TYPE "Sensor Check Struct"
VERSION : 0.1


  STRUCT
   Rising_Pulse_1 : BOOL ;
   Rising_Pulse_2 : BOOL ;
   Memory_Bit_1 : BOOL ;
   Memory_Bit_2 : BOOL ;
   Word_buffer : INT ;
   Word_Result : INT ;
  END_STRUCT ;
END_TYPE

TYPE "CounterCmd"


  STRUCT
   JOB_WR : STRUCT 	// write commands
    NO : BYTE ;	// number
    BUSY : BOOL ;	// job in working
    DONE : BOOL ;	// job is done
    IMPOSS : BOOL ;	// job impossible
    UNKOWN : BOOL ;	// job unkown
   END_STRUCT ;
   JOB_RD : STRUCT 	// read commands
    NO : BYTE ;	// number
    BUSY : BOOL ;	// job in working
    DONE : BOOL ;	// job is done
    IMPOSS : BOOL ;	// job impossible
    UNKOWN : BOOL ;	// job unkown
   END_STRUCT ;
   RESERV_0 : ARRAY  [1 .. 3 ] OF WORD  := 3 (W#16#0) ;	// reserved
   RESERV_1 : WORD ;	// reserved
   MOD_ADR : WORD ;	// module address
   CH_ADR : DWORD ;	// channel address
   DS_OFFS : BYTE ;	// data block offset
   RESERV_2 : BYTE ;	// reserved
   CONTROL_SIGNALS : STRUCT 	// control signals
    BIT0_0 : BOOL ;	// reserved
    BIT0_1 : BOOL ;	// reserved
    BIT0_2 : BOOL ;	// reserved
    BIT0_3 : BOOL ;	// reserved
    BIT0_4 : BOOL ;	// reserved
    BIT0_5 : BOOL ;	// reserved
    BIT0_6 : BOOL ;	// reserved
    BIT0_7 : BOOL ;	// reserved
    CTRL_DQ0 : BOOL ;	// control digital output DQ0
    CTRL_DQ1 : BOOL ;	// control digital output DQ1
    CTRL_DQ2 : BOOL ;	// control digital output DQ2
    CTRL_DQ3 : BOOL ;	// control digital output DQ3
    CTRL_DQ4 : BOOL ;	// control digital output DQ4
    CTRL_DQ5 : BOOL ;	// control digital output DQ5
    CTRL_DQ6 : BOOL ;	// control digital output DQ6
    CTRL_DQ7 : BOOL ;	// control digital output DQ7
    SET_DQ0 : BOOL ;	// set digital output DQ0
    SET_DQ1 : BOOL ;	// set digital output DQ1
    SET_DQ2 : BOOL ;	// set digital output DQ2
    SET_DQ3 : BOOL ;	// set digital output DQ3
    SET_DQ4 : BOOL ;	// set digital output DQ4
    SET_DQ5 : BOOL ;	// set digital output DQ5
    SET_DQ6 : BOOL ;	// set digital output DQ6
    SET_DQ7 : BOOL ;	// set digital output DQ7
    SW_GATE0 : BOOL ;	// software gate 0
    SW_GATE1 : BOOL ;	// software gate 1
    SW_GATE2 : BOOL ;	// software gate 2
    SW_GATE3 : BOOL ;	// software gate 3
    SW_GATE4 : BOOL ;	// software gate 4
    SW_GATE5 : BOOL ;	// software gate 5
    SW_GATE6 : BOOL ;	// software gate 6
    SW_GATE7 : BOOL ;	// software gate 7
    CTRL_DWORD1 : DWORD ;	// reserved
    CTRL_DWORD2 : DWORD ;	// reserved
    CTRL_DWORD3 : DWORD ;	// reserved
   END_STRUCT ;
   CHECKBACK_SIGNALS : STRUCT 	// checkback signals
    BIT0_0 : BOOL ;	// reserved
    STS_TFB : BOOL ;	// status test free bit
    BIT0_2 : BOOL ;	// reserved
    BIT0_3 : BOOL ;	// reserved
    DATA_ERR : BOOL ;	// data error bit
    BIT0_5 : BOOL ;	// reserved
    BIT0_6 : BOOL ;	// reserved
    PARA : BOOL ;	// module parametrized
    STS_CMP0 : BOOL ;	// status compare event 0
    STS_CMP1 : BOOL ;	// status compare event 1
    STS_CMP2 : BOOL ;	// status compare event 2
    STS_CMP3 : BOOL ;	// status compare event 3
    STS_CMP4 : BOOL ;	// status compare event 4
    STS_CMP5 : BOOL ;	// status compare event 5
    STS_CMP6 : BOOL ;	// status compare event 6
    STS_CMP7 : BOOL ;	// status compare event 7
    STS_UFLW0 : BOOL ;	// status counter 0 passed the underflow value
    STS_UFLW1 : BOOL ;	// status counter 1 passed the underflow value
    STS_UFLW2 : BOOL ;	// status counter 2 passed the underflow value
    STS_UFLW3 : BOOL ;	// status counter 3 passed the underflow value
    STS_UFLW4 : BOOL ;	// status counter 4 passed the underflow value
    STS_UFLW5 : BOOL ;	// status counter 5 passed the underflow value
    STS_UFLW6 : BOOL ;	// status counter 6 passed the underflow value
    STS_UFLW7 : BOOL ;	// status counter 7 passed the underflow value
    STS_OFLW0 : BOOL ;	// status counter 0 passed the overflow value
    STS_OFLW1 : BOOL ;	// status counter 1 passed the overflow value
    STS_OFLW2 : BOOL ;	// status counter 2 passed the overflow value
    STS_OFLW3 : BOOL ;	// status counter 3 passed the overflow value
    STS_OFLW4 : BOOL ;	// status counter 4 passed the overflow value
    STS_OFLW5 : BOOL ;	// status counter 5 passed the overflow value
    STS_OFLW6 : BOOL ;	// status counter 6 passed the overflow value
    STS_OFLW7 : BOOL ;	// status counter 7 passed the overflow value
    STS_DIR0 : BOOL ;	// status counter 0 direction
    STS_DIR1 : BOOL ;	// status counter 1 direction
    STS_DIR2 : BOOL ;	// status counter 2 direction
    STS_DIR3 : BOOL ;	// status counter 3 direction
    STS_DIR4 : BOOL ;	// status counter 4 direction
    STS_DIR5 : BOOL ;	// status counter 5 direction
    STS_DIR6 : BOOL ;	// status counter 6 direction
    STS_DIR7 : BOOL ;	// status counter 7 direction
    STS_DI0 : BOOL ;	// status of the digital input 0
    STS_DI1 : BOOL ;	// status of the digital input 1
    STS_DI2 : BOOL ;	// status of the digital input 2
    STS_DI3 : BOOL ;	// status of the digital input 3
    STS_DI4 : BOOL ;	// status of the digital input 4
    STS_DI5 : BOOL ;	// status of the digital input 5
    STS_DI6 : BOOL ;	// status of the digital input 6
    STS_DI7 : BOOL ;	// status of the digital input 7
    STS_DQ0 : BOOL ;	// status of the digital output 0
    STS_DQ1 : BOOL ;	// status of the digital output 1
    STS_DQ2 : BOOL ;	// status of the digital output 2
    STS_DQ3 : BOOL ;	// status of the digital output 3
    STS_DQ4 : BOOL ;	// status of the digital output 4
    STS_DQ5 : BOOL ;	// status of the digital output 5
    STS_DQ6 : BOOL ;	// status of the digital output 6
    STS_DQ7 : BOOL ;	// status of the digital output 7
    STS_GATE0 : BOOL ;	// status of the internal gate 0
    STS_GATE1 : BOOL ;	// status of the internal gate 1
    STS_GATE2 : BOOL ;	// status of the internal gate 2
    STS_GATE3 : BOOL ;	// status of the internal gate 3
    STS_GATE4 : BOOL ;	// status of the internal gate 4
    STS_GATE5 : BOOL ;	// status of the internal gate 5
    STS_GATE6 : BOOL ;	// status of the internal gate 6
    STS_GATE7 : BOOL ;	// status of the internal gate 7
    USER_STAT_WORD0 : WORD ;	// user specific status
    USER_STAT_WORD1 : WORD ;	// user specific status
    USER_STAT_WORD2 : WORD ;	// user specific status
    USER_STAT_WORD3 : WORD ;	// user specific status
   END_STRUCT ;
   LOAD_VAL0 : DINT ;	// load value counter 0
   LOAD_VAL1 : DINT ;	// load value counter 1
   LOAD_VAL2 : DINT ;	// load value counter 2
   LOAD_VAL3 : DINT ;	// load value counter 3
   LOAD_VAL4 : DINT ;	// load value counter 4
   LOAD_VAL5 : DINT ;	// load value counter 5
   LOAD_VAL6 : DINT ;	// load value counter 6
   LOAD_VAL7 : DINT ;	// load value counter 7
   LOAD_PREPARE_VAL0 : DINT ;	// load prepare value counter 0
   LOAD_PREPARE_VAL1 : DINT ;	// load prepare value counter 1
   LOAD_PREPARE_VAL2 : DINT ;	// load prepare value counter 2
   LOAD_PREPARE_VAL3 : DINT ;	// load prepare value counter 3
   LOAD_PREPARE_VAL4 : DINT ;	// load prepare value counter 4
   LOAD_PREPARE_VAL5 : DINT ;	// load prepare value counter 5
   LOAD_PREPARE_VAL6 : DINT ;	// load prepare value counter 6
   LOAD_PREPARE_VAL7 : DINT ;	// load prepare value counter 7
   CMP_VAL0 : DINT ;	// comparator value 0
   CMP_VAL1 : DINT ;	// comparator value 1
   CMP_VAL2 : DINT ;	// comparator value 2
   CMP_VAL3 : DINT ;	// comparator value 3
   CMP_VAL4 : DINT ;	// comparator value 4
   CMP_VAL5 : DINT ;	// comparator value 5
   CMP_VAL6 : DINT ;	// comparator value 6
   CMP_VAL7 : DINT ;	// comparator value 7
   ACT_CNTV0 : DINT ;	// actual counter value 0
   ACT_MSRV0 : DINT ;	// act. measurement value 0
   ACT_CNTV1 : DINT ;	// actual counter value 1
   ACT_MSRV1 : DINT ;	// act. measurement value 1
   ACT_CNTV2 : DINT ;	// actual counter value 2
   ACT_MSRV2 : DINT ;	// act. measurement value 2
   ACT_CNTV3 : DINT ;	// actual counter value 3
   ACT_MSRV3 : DINT ;	// act. measurement value 3
   ACT_CNTV4 : DINT ;	// actual counter value 4
   ACT_MSRV4 : DINT ;	// act. measurement value 4
   ACT_CNTV5 : DINT ;	// actual counter value 5
   ACT_MSRV5 : DINT ;	// act. measurement value 5
   ACT_CNTV6 : DINT ;	// actual counter value 6
   ACT_MSRV6 : DINT ;	// act. measurement value 6
   ACT_CNTV7 : DINT ;	// actual counter value 7
   ACT_MSRV7 : DINT ;	// act. measurement value 7
   DIAGNOSTIC_INT_INFO : STRUCT 	// diagnostic int. information
    BYTE0 : BYTE ;	// byte 0
    BYTE1 : BYTE ;	// byte 1
    BYTE2 : BYTE ;	// byte 2
    BYTE3 : BYTE ;	// byte 3
    BYTE4 : BYTE ;	// channel type info
    BYTE5 : BYTE ;	// channel info length
    BYTE6 : BYTE ;	// number of channels
    BYTE7 : BYTE ;	// channel error vector
    BYTE8 : BYTE ;	// error counter 0
    BYTE9 : BYTE ;	// error counter 1
    BYTE10 : BYTE ;	// error counter 2
    BYTE11 : BYTE ;	// error counter 3
    BYTE12 : BYTE ;	// error counter 4
    BYTE13 : BYTE ;	// error counter 5
    BYTE14 : BYTE ;	// error counter 6
    BYTE15 : BYTE ;	// error counter 7
   END_STRUCT ;
  END_STRUCT ;
END_TYPE

TYPE "Sensor Debounce Struct"
VERSION : 0.1


  STRUCT
   Rising_Pulse_1 : BOOL ;
   Rising_Pulse_2 : BOOL ;
   Rising_Pulse_3 : BOOL ;
   Rising_Pulse_4 : BOOL ;
   Rising_Pulse_5 : BOOL ;
   Rising_Pulse_6 : BOOL ;
   Rising_Pulse_7 : BOOL ;
   Rising_Pulse_8 : BOOL ;
   Bit_0_FrontEnd : BOOL ;
   Bit_1_FrontEnd : BOOL ;
   Bit_0_RearEnd : BOOL ;
   Bit_1_RearEnd : BOOL ;
   Packet_Exiting : BOOL ;
   Count_Error : BOOL ;
   Sens_Error : BOOL ;
   FirstScan_Init_Done : BOOL ;
   Bit_0_ON_Time : INT ;	//Count Up Sens
   Bit_1_ON_Time : INT ;	//Count Dn Sens
   Word_Count_Result : INT ;
   Word_Count_Limit : INT ;
  END_STRUCT ;
END_TYPE

TYPE "Sensor U Shape Struct"
VERSION : 0.1


  STRUCT
   RISING_PULSE_1 : BOOL ;
   RISING_PULSE_2 : BOOL ;
   RISING_PULSE_3 : BOOL ;
   RISING_PULSE_4 : BOOL ;
   RISING_PULSE_5 : BOOL ;
   RISING_PULSE_6 : BOOL ;
   RISING_PULSE_7 : BOOL ;
   RISING_PULSE_8 : BOOL ;
   EVT_ACTIVE_0 : BOOL ;
   EVT_VALIDATED_0 : BOOL ;
   EVT_REJECTED_0 : BOOL ;
   EVT_ACTIVE_1 : BOOL ;
   BYPASS_LONG_0 : BOOL ;
   INIT_DONE : BOOL ;
   SPARE_1 : BOOL ;
   SPARE_2 : BOOL ;
   TMR_0_mS : INT ;
   TMR_1_mS : INT ;
   RESULT_SHORT_0 : INT ;
   VALIDATE_0_mS : INT ;
   DEBOUNCE_1_mS : INT ;
   COUNT_LIMIT : INT ;
  END_STRUCT ;
END_TYPE

TYPE "Debouncer Counter Struct"
VERSION : 0.7


  STRUCT
   FirstScan_Done : BOOL ;	//Init Done
   Bit0_ON_Latch : BOOL ;	//InFeed - Packet Seen (Until Gap)
   Bit1_ON_Latch : BOOL ;	//Exit - Packet Seen During Transfer (Until Gap)
   Transfer_Active : BOOL ;	//Spare (Compatibility)
   Count_Done_Latch_0 : BOOL ;	//InFeed - Packet Counted
   Count_Done_Latch_1 : BOOL ;	//Spare (Compatibility)
   Error : BOOL ;	//InFeed Sensor Stuck
   Spare_Bit : BOOL ;	//Spare
   Bit0_Entry_mS : INT ;	//InFeed - ON Time This Packet [mS]
   Bit0_OFF_mS : INT ;	//InFeed - Gap Time [mS]
   Bit0_Stuck_mS : INT ;	//InFeed - Continuous ON Time [mS]
   Bit1_Exit_mS : INT ;	//Exit - ON Time During Transfer [mS]
   Bit1_OFF_mS : INT ;	//Exit - Gap Time [mS]
   Space_Between : INT ;	//Gap Confirm [mS]
   InFeed_Window_mS : INT ;	//Info: Preset Used [mS]
   Exit_Window_mS : INT ;	//Butted Packets Window [mS]
   Count_Result : INT ;	//Packet Count
   Maximum_Count : INT ;	//Count Limit (0 = No Limit)
   HMI_Last : INT ;	//Last Value Written to HMI
  END_STRUCT ;
END_TYPE

TYPE "Width Sensor Struct"
VERSION : 0.9


  STRUCT
   Was_On : BOOL ;	//Sensor State Last Scan
   Open : BOOL ;	//Packet in Progress
   Low : BOOL ;	//Sensor OFF Inside a Packet (Sag or Gap - Not Decided Yet)
   Skip : BOOL ;	//Packet Already Covering at Start = Partial, Not Recorded
   Front : BOOL ;	//New Packet Front This Scan (Pulse)
   Spare_2 : BOOL ;
   Spare_3 : BOOL ;
   Spare_4 : BOOL ;
   Start_Pos : DINT ;	//Encoder at Packet Front [Pulses]
   Fall_Pos : DINT ;	//Encoder at Last OFF [Pulses]
   Count : INT ;	//Packets Measured This Transfer
   Skipped : INT ;	//Partial Packets Not Measured (0 or 1)
   Sag_Count : INT ;	//OFF Shorter than Gap_Min = Sag (U-Shape / Low Packet)
   Width_Sum_mm : DINT ;	//Sum of Widths [mm]
   Width_Min_mm : INT ;	//Smallest Width [mm]
   Width_Max_mm : INT ;	//Largest Width [mm]
   Width_Avg_mm : INT ;	//Average Width [mm]
   Last_Width_mm : INT ;	//Last Packet Width [mm]
   Sag_Max_mm : INT ;	//Longest Sag [mm]
   Gap_Min_mm : INT ;	//Shortest Real Gap Between Packets [mm]
   Time_ms : DINT ;	//Time Since Packet Front [mS]
   Fall_ms : DINT ;	//Time at Last OFF [mS]
   Width_Sum_ms : DINT ;	//Sum of Widths [mS]
   Width_Avg_ms : INT ;	//Average Width [mS] @ C10 Fast = C11/C12/C21/C22 Speed
   Last_Width_ms : INT ;	//Last Packet Width [mS]
  END_STRUCT ;
END_TYPE

TYPE "Blanking Struct"
VERSION : 0.1


  STRUCT
   Was_On : BOOL ;	//Sensor State Last Scan
   Pulse : BOOL ;	//Cleaned Packet Pulse (Info)
   Spare_1 : BOOL ;
   Spare_2 : BOOL ;
   Spare_3 : BOOL ;
   Spare_4 : BOOL ;
   Spare_5 : BOOL ;
   Spare_6 : BOOL ;
   T_ms : DINT  := L#60000;	//Belt Run Time Since Last Counted Packet [mS]
   Pulse_ms : INT ;	//Pulse Time Left [mS]
   Count : INT ;	//Packets Counted (Cleaned) - Total
   Raw : INT ;	//Raw Sensor Fronts - Total
   Sag : INT ;	//Fronts Ignored (Inside Blanking = Sag of a U-Shape) - Total
   Butt : INT ;	//Butted Packets Counted (Sensor Never Cleared) - Total
  END_STRUCT ;
END_TYPE

DATA_BLOCK "DB UTILITY"
TITLE =
VERSION : 0.1


  STRUCT
   DB_VAR : INT ;	//Temporary placeholder variable
   VAL_TMP_SEC_MS_PCS : INT ;	//Temporary placeholder variable
   RAZ_TMR_RESTART_PCS : BOOL ;	// PCS
   VAL_CMP_RESTART_PCS_OS : BOOL ;	// PCS
   VAL_CMP_RESTART_PCS : BOOL ;
   DEM_RESTART_PCS : BOOL ;
   DB_bool4 : BOOL ;	//Temporary placeholder variable
   DB_bool5 : BOOL ;	//Temporary placeholder variable
   DB_bool6 : BOOL ;	//Temporary placeholder variable
   DB_bool7 : BOOL ;	//Temporary placeholder variable
   DB_bool8 : BOOL ;	//Temporary placeholder variable
   DB_bool9 : BOOL ;	//Temporary placeholder variable
   DB_bool10 : BOOL ;	//Temporary placeholder variable
   DB_bool11 : BOOL ;	//Temporary placeholder variable
   DB_bool12 : BOOL ;	//Temporary placeholder variable
   DB_bool13 : BOOL ;	//Temporary placeholder variable
   DB_bool14 : BOOL ;	//Temporary placeholder variable
   C4_Moving : BOOL ;	//Conveyor 4 is Moving
   Scan_Cycle_Previous : INT ;	//Previous Scan Cycle - OB1
   DB_VAR4 : INT ;	//Temporary placeholder variable
   LENGTH_CONST : REAL ;	//Packet Constant - Length
   WIDTH_CONST : REAL ;	//Packet Constant - Width
   DB_VAR7 : INT ;	//Temporary placeholder variable
   Pusher_0_Disable : BOOL ;	//Pusher 0 Disable
   Elevator_Disable : BOOL ;	//Elevator Disable
   Pusher_1_Disable : BOOL ;	//Pusher 1 Disable
   Conveyor_1_Disable : BOOL ;	//Conveyor 1 Disable
   Conveyor_2_Disable : BOOL ;	//Conveyor 2 Disable
   Conveyor_3_Disable : BOOL ;	//Conveyor 3 Disable
   Conveyor_4_Disable : BOOL ;	//Conveyor 4 Disable
   Conveyor_5_Disable : BOOL ;	//Conveyor 5 Disable
   Conveyor_6_Disable : BOOL ;	//Conveyor 6 Disable
   Conveyor_7_Disable : BOOL ;	//Conveyor 7 Disable
   Conveyor_8_Disable : BOOL ;	//Conveyor 8 Disable
   Conveyor_9_Disable : BOOL ;	//Conveyor 9 Disable
   Pusher_2_Disable : BOOL ;	//Pusher 2 Disable
   Conveyor_10_Disable : BOOL ;	//Conveyor 10 Disable
   Pivot_Disable : BOOL ;	//Pivot Disable
   Conveyor_11_Disable : BOOL ;	//Conveyor 11 Disable
   Conveyor_12_Disable : BOOL ;	//Conveyor 12 Disable
   Conveyor_13_Disable : BOOL ;	//Conveyor 13 Disable
   Conveyor_21_Disable : BOOL ;	//Conveyor 21 Disable
   Conveyor_22_Disable : BOOL ;	//Conveyor 22 Disable
   Conveyor_23_Disable : BOOL ;	//Conveyor 23 Disable
   Feeder_Lift_disable : BOOL ;	//Feeder Lift Disable
   Feeder_Fingers_disable : BOOL ;	//Feeder Fingers Disable
   RESERVE : BOOL ;
   Freeze_Sequence_1 : BOOL ;	//Sequence Freezer Bit - Elevator
   T15_DN : BOOL ;	//Adder Done Elevator 1 Timeout Done
   T19_DN : BOOL ;	//Adder Done Conveyor 1 Timeout Done
   T23_DN : BOOL ;	//Adder Done Conveyor 2 Lift Fault
   T24_DN : BOOL ;	//Adder Done Conveyor 2 Belt Timeout
   T25_DN : BOOL ;	//Adder Done Conveyor 2 Roller Timeout
   T27_DN : BOOL ;	//Adder Done Conveyor 3 Slat Start Pulse 100mS
   T28_DN : BOOL ;	//Adder Done Conveyor 3 Slat Timeout 11s
   T29_DN : BOOL ;	//Adder Done Conveyor 4 LB obstruction alarm 10s
   T90_DN : BOOL ;	//Adder Done Conveyor 4 Encoder-stop helper timers 500ms
   T91_DN : BOOL ;	//Adder Done Conveyor 4 Encoder-stop helper timers 500ms
   T31_DN : BOOL ;	//Adder Done Conveyor 4 InFeed timeout 5s
   T32_DN : BOOL ;	//Adder Done Conveyor 4 Transfer max time 20s
   T33_DN : BOOL ;	//Adder Done Conveyor 4 Clearing timeout 20s
   T35_DN : BOOL ;	//Adder Done Conveyor 5 Link timeout 20s
   Freeze_Sequence_2 : BOOL ;	//Sequence Freezer Bit - Collator
   T15_ET : DINT ;	//Adder Count Elevator 1 Timeout Count 100mS
   T19_ET : DINT ;	//Adder Count Conveyor 1 Timeout Count 10s
   T23_ET : DINT ;	//Adder Count Conveyor 2 Lift Fault TimeOut 2s
   T24_ET : DINT ;	//Adder Count Conveyor 2 Belt Timeout 2.5s
   T25_ET : DINT ;	//Adder Count Conveyor 2 Roller Extended RunTime 8s
   T27_ET : DINT ;	//Adder Count Conveyor 3 Slat Start Pulse 100mS
   T28_ET : DINT ;	//Adder Count Conveyor 3 Slat Timeout 11s
   T29_ET : DINT ;	//Adder Count Conveyor 4 LB obstruction alarm 10s
   T90_ET : DINT ;	//Adder Count Conveyor 4 Encoder-stop helper timers 500ms
   T91_ET : DINT ;	//Adder Count Conveyor 4 Encoder-stop helper timers 500ms
   T31_ET : DINT ;	//Adder Count Conveyor 4 InFeed timeout 5s
   T32_ET : DINT ;	//Adder Count Conveyor 4 Transfer max time 20s
   T33_ET : DINT ;	//Adder Count Conveyor 4 Clearing timeout 20s
   T35_ET : DINT ;	//Adder Count Conveyor 5 Link timeout 20s
  END_STRUCT ;
BEGIN
   DB_VAR := 0;
   VAL_TMP_SEC_MS_PCS := 13886;
   RAZ_TMR_RESTART_PCS := FALSE;
   VAL_CMP_RESTART_PCS_OS := FALSE;
   VAL_CMP_RESTART_PCS := FALSE;
   DEM_RESTART_PCS := FALSE;
   DB_bool4 := FALSE;
   DB_bool5 := FALSE;
   DB_bool6 := FALSE;
   DB_bool7 := FALSE;
   DB_bool8 := FALSE;
   DB_bool9 := FALSE;
   DB_bool10 := FALSE;
   DB_bool11 := FALSE;
   DB_bool12 := FALSE;
   DB_bool13 := FALSE;
   DB_bool14 := FALSE;
   C4_Moving := FALSE;
   Scan_Cycle_Previous := 8;
   DB_VAR4 := 0;
   LENGTH_CONST := 0.000000e+000;
   WIDTH_CONST := 0.000000e+000;
   DB_VAR7 := 0;
   Pusher_0_Disable := FALSE;
   Elevator_Disable := FALSE;
   Pusher_1_Disable := FALSE;
   Conveyor_1_Disable := FALSE;
   Conveyor_2_Disable := FALSE;
   Conveyor_3_Disable := FALSE;
   Conveyor_4_Disable := FALSE;
   Conveyor_5_Disable := FALSE;
   Conveyor_6_Disable := FALSE;
   Conveyor_7_Disable := FALSE;
   Conveyor_8_Disable := FALSE;
   Conveyor_9_Disable := FALSE;
   Pusher_2_Disable := FALSE;
   Conveyor_10_Disable := FALSE;
   Pivot_Disable := FALSE;
   Conveyor_11_Disable := FALSE;
   Conveyor_12_Disable := FALSE;
   Conveyor_13_Disable := FALSE;
   Conveyor_21_Disable := FALSE;
   Conveyor_22_Disable := FALSE;
   Conveyor_23_Disable := FALSE;
   Feeder_Lift_disable := FALSE;
   Feeder_Fingers_disable := FALSE;
   RESERVE := FALSE;
   Freeze_Sequence_1 := FALSE;
   T15_DN := FALSE;
   T19_DN := FALSE;
   T23_DN := FALSE;
   T24_DN := FALSE;
   T25_DN := FALSE;
   T27_DN := FALSE;
   T28_DN := FALSE;
   T29_DN := FALSE;
   T90_DN := FALSE;
   T91_DN := FALSE;
   T31_DN := FALSE;
   T32_DN := FALSE;
   T33_DN := FALSE;
   T35_DN := FALSE;
   Freeze_Sequence_2 := FALSE;
   T15_ET := L#0;
   T19_ET := L#0;
   T23_ET := L#0;
   T24_ET := L#0;
   T25_ET := L#0;
   T27_ET := L#0;
   T28_ET := L#0;
   T29_ET := L#0;
   T90_ET := L#0;
   T91_ET := L#0;
   T31_ET := L#0;
   T32_ET := L#0;
   T33_ET := L#0;
   T35_ET := L#0;
END_DATA_BLOCK

DATA_BLOCK "FM350 DB"
TITLE =
VERSION : 0.1

"CounterCmd"
BEGIN
   JOB_WR.NO := B#16#0;
   JOB_WR.BUSY := FALSE;
   JOB_WR.DONE := FALSE;
   JOB_WR.IMPOSS := FALSE;
   JOB_WR.UNKOWN := FALSE;
   JOB_RD.NO := B#16#0;
   JOB_RD.BUSY := FALSE;
   JOB_RD.DONE := FALSE;
   JOB_RD.IMPOSS := FALSE;
   JOB_RD.UNKOWN := FALSE;
   RESERV_0[1] := W#16#0;
   RESERV_0[2] := W#16#0;
   RESERV_0[3] := W#16#0;
   RESERV_1 := W#16#0;
   MOD_ADR := W#16#0;
   CH_ADR := DW#16#0;
   DS_OFFS := B#16#0;
   RESERV_2 := B#16#0;
   CONTROL_SIGNALS.BIT0_0 := FALSE;
   CONTROL_SIGNALS.BIT0_1 := FALSE;
   CONTROL_SIGNALS.BIT0_2 := FALSE;
   CONTROL_SIGNALS.BIT0_3 := FALSE;
   CONTROL_SIGNALS.BIT0_4 := FALSE;
   CONTROL_SIGNALS.BIT0_5 := FALSE;
   CONTROL_SIGNALS.BIT0_6 := FALSE;
   CONTROL_SIGNALS.BIT0_7 := FALSE;
   CONTROL_SIGNALS.CTRL_DQ0 := FALSE;
   CONTROL_SIGNALS.CTRL_DQ1 := FALSE;
   CONTROL_SIGNALS.CTRL_DQ2 := FALSE;
   CONTROL_SIGNALS.CTRL_DQ3 := FALSE;
   CONTROL_SIGNALS.CTRL_DQ4 := FALSE;
   CONTROL_SIGNALS.CTRL_DQ5 := FALSE;
   CONTROL_SIGNALS.CTRL_DQ6 := FALSE;
   CONTROL_SIGNALS.CTRL_DQ7 := FALSE;
   CONTROL_SIGNALS.SET_DQ0 := FALSE;
   CONTROL_SIGNALS.SET_DQ1 := FALSE;
   CONTROL_SIGNALS.SET_DQ2 := FALSE;
   CONTROL_SIGNALS.SET_DQ3 := FALSE;
   CONTROL_SIGNALS.SET_DQ4 := FALSE;
   CONTROL_SIGNALS.SET_DQ5 := FALSE;
   CONTROL_SIGNALS.SET_DQ6 := FALSE;
   CONTROL_SIGNALS.SET_DQ7 := FALSE;
   CONTROL_SIGNALS.SW_GATE0 := FALSE;
   CONTROL_SIGNALS.SW_GATE1 := FALSE;
   CONTROL_SIGNALS.SW_GATE2 := FALSE;
   CONTROL_SIGNALS.SW_GATE3 := FALSE;
   CONTROL_SIGNALS.SW_GATE4 := FALSE;
   CONTROL_SIGNALS.SW_GATE5 := FALSE;
   CONTROL_SIGNALS.SW_GATE6 := FALSE;
   CONTROL_SIGNALS.SW_GATE7 := FALSE;
   CONTROL_SIGNALS.CTRL_DWORD1 := DW#16#0;
   CONTROL_SIGNALS.CTRL_DWORD2 := DW#16#0;
   CONTROL_SIGNALS.CTRL_DWORD3 := DW#16#0;
   CHECKBACK_SIGNALS.BIT0_0 := FALSE;
   CHECKBACK_SIGNALS.STS_TFB := FALSE;
   CHECKBACK_SIGNALS.BIT0_2 := FALSE;
   CHECKBACK_SIGNALS.BIT0_3 := FALSE;
   CHECKBACK_SIGNALS.DATA_ERR := FALSE;
   CHECKBACK_SIGNALS.BIT0_5 := FALSE;
   CHECKBACK_SIGNALS.BIT0_6 := FALSE;
   CHECKBACK_SIGNALS.PARA := FALSE;
   CHECKBACK_SIGNALS.STS_CMP0 := FALSE;
   CHECKBACK_SIGNALS.STS_CMP1 := FALSE;
   CHECKBACK_SIGNALS.STS_CMP2 := FALSE;
   CHECKBACK_SIGNALS.STS_CMP3 := FALSE;
   CHECKBACK_SIGNALS.STS_CMP4 := FALSE;
   CHECKBACK_SIGNALS.STS_CMP5 := FALSE;
   CHECKBACK_SIGNALS.STS_CMP6 := FALSE;
   CHECKBACK_SIGNALS.STS_CMP7 := FALSE;
   CHECKBACK_SIGNALS.STS_UFLW0 := FALSE;
   CHECKBACK_SIGNALS.STS_UFLW1 := FALSE;
   CHECKBACK_SIGNALS.STS_UFLW2 := FALSE;
   CHECKBACK_SIGNALS.STS_UFLW3 := FALSE;
   CHECKBACK_SIGNALS.STS_UFLW4 := FALSE;
   CHECKBACK_SIGNALS.STS_UFLW5 := FALSE;
   CHECKBACK_SIGNALS.STS_UFLW6 := FALSE;
   CHECKBACK_SIGNALS.STS_UFLW7 := FALSE;
   CHECKBACK_SIGNALS.STS_OFLW0 := FALSE;
   CHECKBACK_SIGNALS.STS_OFLW1 := FALSE;
   CHECKBACK_SIGNALS.STS_OFLW2 := FALSE;
   CHECKBACK_SIGNALS.STS_OFLW3 := FALSE;
   CHECKBACK_SIGNALS.STS_OFLW4 := FALSE;
   CHECKBACK_SIGNALS.STS_OFLW5 := FALSE;
   CHECKBACK_SIGNALS.STS_OFLW6 := FALSE;
   CHECKBACK_SIGNALS.STS_OFLW7 := FALSE;
   CHECKBACK_SIGNALS.STS_DIR0 := FALSE;
   CHECKBACK_SIGNALS.STS_DIR1 := FALSE;
   CHECKBACK_SIGNALS.STS_DIR2 := FALSE;
   CHECKBACK_SIGNALS.STS_DIR3 := FALSE;
   CHECKBACK_SIGNALS.STS_DIR4 := FALSE;
   CHECKBACK_SIGNALS.STS_DIR5 := FALSE;
   CHECKBACK_SIGNALS.STS_DIR6 := FALSE;
   CHECKBACK_SIGNALS.STS_DIR7 := FALSE;
   CHECKBACK_SIGNALS.STS_DI0 := FALSE;
   CHECKBACK_SIGNALS.STS_DI1 := FALSE;
   CHECKBACK_SIGNALS.STS_DI2 := FALSE;
   CHECKBACK_SIGNALS.STS_DI3 := FALSE;
   CHECKBACK_SIGNALS.STS_DI4 := FALSE;
   CHECKBACK_SIGNALS.STS_DI5 := FALSE;
   CHECKBACK_SIGNALS.STS_DI6 := FALSE;
   CHECKBACK_SIGNALS.STS_DI7 := FALSE;
   CHECKBACK_SIGNALS.STS_DQ0 := FALSE;
   CHECKBACK_SIGNALS.STS_DQ1 := FALSE;
   CHECKBACK_SIGNALS.STS_DQ2 := FALSE;
   CHECKBACK_SIGNALS.STS_DQ3 := FALSE;
   CHECKBACK_SIGNALS.STS_DQ4 := FALSE;
   CHECKBACK_SIGNALS.STS_DQ5 := FALSE;
   CHECKBACK_SIGNALS.STS_DQ6 := FALSE;
   CHECKBACK_SIGNALS.STS_DQ7 := FALSE;
   CHECKBACK_SIGNALS.STS_GATE0 := FALSE;
   CHECKBACK_SIGNALS.STS_GATE1 := FALSE;
   CHECKBACK_SIGNALS.STS_GATE2 := FALSE;
   CHECKBACK_SIGNALS.STS_GATE3 := FALSE;
   CHECKBACK_SIGNALS.STS_GATE4 := FALSE;
   CHECKBACK_SIGNALS.STS_GATE5 := FALSE;
   CHECKBACK_SIGNALS.STS_GATE6 := FALSE;
   CHECKBACK_SIGNALS.STS_GATE7 := FALSE;
   CHECKBACK_SIGNALS.USER_STAT_WORD0 := W#16#0;
   CHECKBACK_SIGNALS.USER_STAT_WORD1 := W#16#0;
   CHECKBACK_SIGNALS.USER_STAT_WORD2 := W#16#0;
   CHECKBACK_SIGNALS.USER_STAT_WORD3 := W#16#0;
   LOAD_VAL0 := L#0;
   LOAD_VAL1 := L#0;
   LOAD_VAL2 := L#0;
   LOAD_VAL3 := L#0;
   LOAD_VAL4 := L#0;
   LOAD_VAL5 := L#0;
   LOAD_VAL6 := L#0;
   LOAD_VAL7 := L#0;
   LOAD_PREPARE_VAL0 := L#0;
   LOAD_PREPARE_VAL1 := L#0;
   LOAD_PREPARE_VAL2 := L#0;
   LOAD_PREPARE_VAL3 := L#0;
   LOAD_PREPARE_VAL4 := L#0;
   LOAD_PREPARE_VAL5 := L#0;
   LOAD_PREPARE_VAL6 := L#0;
   LOAD_PREPARE_VAL7 := L#0;
   CMP_VAL0 := L#0;
   CMP_VAL1 := L#0;
   CMP_VAL2 := L#0;
   CMP_VAL3 := L#0;
   CMP_VAL4 := L#0;
   CMP_VAL5 := L#0;
   CMP_VAL6 := L#0;
   CMP_VAL7 := L#0;
   ACT_CNTV0 := L#0;
   ACT_MSRV0 := L#0;
   ACT_CNTV1 := L#0;
   ACT_MSRV1 := L#0;
   ACT_CNTV2 := L#0;
   ACT_MSRV2 := L#0;
   ACT_CNTV3 := L#0;
   ACT_MSRV3 := L#0;
   ACT_CNTV4 := L#0;
   ACT_MSRV4 := L#0;
   ACT_CNTV5 := L#0;
   ACT_MSRV5 := L#0;
   ACT_CNTV6 := L#0;
   ACT_MSRV6 := L#0;
   ACT_CNTV7 := L#0;
   ACT_MSRV7 := L#0;
   DIAGNOSTIC_INT_INFO.BYTE0 := B#16#0;
   DIAGNOSTIC_INT_INFO.BYTE1 := B#16#0;
   DIAGNOSTIC_INT_INFO.BYTE2 := B#16#0;
   DIAGNOSTIC_INT_INFO.BYTE3 := B#16#0;
   DIAGNOSTIC_INT_INFO.BYTE4 := B#16#0;
   DIAGNOSTIC_INT_INFO.BYTE5 := B#16#0;
   DIAGNOSTIC_INT_INFO.BYTE6 := B#16#0;
   DIAGNOSTIC_INT_INFO.BYTE7 := B#16#0;
   DIAGNOSTIC_INT_INFO.BYTE8 := B#16#0;
   DIAGNOSTIC_INT_INFO.BYTE9 := B#16#0;
   DIAGNOSTIC_INT_INFO.BYTE10 := B#16#0;
   DIAGNOSTIC_INT_INFO.BYTE11 := B#16#0;
   DIAGNOSTIC_INT_INFO.BYTE12 := B#16#0;
   DIAGNOSTIC_INT_INFO.BYTE13 := B#16#0;
   DIAGNOSTIC_INT_INFO.BYTE14 := B#16#0;
   DIAGNOSTIC_INT_INFO.BYTE15 := B#16#0;
END_DATA_BLOCK

DATA_BLOCK "DB SENSOR CHECK"
TITLE =
VERSION : 0.1


  STRUCT
   B5_1 : "Sensor Check Struct";
   B5_2 : "Sensor Check Struct";
   B5_4 : "Sensor Check Struct";
   B5_5 : "Sensor Check Struct";
   B6_0 : "Sensor Check Struct";
   B6_1 : "Sensor Check Struct";
   B6_2 : "Sensor Check Struct";
   B6_4 : "Sensor Check Struct";
   B6_7 : "Sensor Check Struct";
   B7_0 : "Sensor Check Struct";
   B7_1 : "Sensor Check Struct";
   B7_2 : "Sensor Check Struct";
   B7_3 : "Sensor Check Struct";
   B7_4 : "Sensor Check Struct";
   B8_2 : "Sensor Check Struct";
   B9_6 : "Sensor Check Struct";
   B9_7 : "Sensor Check Struct";
   B10_3 : "Sensor Check Struct";
   B10_4 : "Sensor Check Struct";
   B10_5 : "Sensor Check Struct";
   B10_6 : "Sensor Check Struct";
   B10_7 : "Sensor Check Struct";
   B11_0 : "Sensor Check Struct";
   B11_1 : "Sensor Check Struct";
   B12_3 : "Sensor Check Struct";
   B13_0 : "Sensor Check Struct";
   B15_4 : "Sensor Check Struct";
   B15_5 : "Sensor Check Struct";
   B15_6 : "Sensor Check Struct";
   B15_7 : "Sensor Check Struct";
   B35_2 : "Sensor Check Struct";
   B35_3 : "Sensor Check Struct";
   B35_4 : "Sensor Check Struct";
   B11_2 : "Sensor Check Struct";
   Z2040 : BOOL ;
   M052 : BOOL ;
   M1122 : BOOL ;
   M1123 : BOOL ;
   M1124 : BOOL ;
   M1125 : BOOL ;
   M1126 : BOOL ;
   M1127 : BOOL ;
  END_STRUCT ;
BEGIN
   B5_1.Rising_Pulse_1 := FALSE;
   B5_1.Rising_Pulse_2 := FALSE;
   B5_1.Memory_Bit_1 := FALSE;
   B5_1.Memory_Bit_2 := FALSE;
   B5_1.Word_buffer := 0;
   B5_1.Word_Result := 0;
   B5_2.Rising_Pulse_1 := FALSE;
   B5_2.Rising_Pulse_2 := FALSE;
   B5_2.Memory_Bit_1 := FALSE;
   B5_2.Memory_Bit_2 := FALSE;
   B5_2.Word_buffer := 0;
   B5_2.Word_Result := 0;
   B5_4.Rising_Pulse_1 := FALSE;
   B5_4.Rising_Pulse_2 := FALSE;
   B5_4.Memory_Bit_1 := FALSE;
   B5_4.Memory_Bit_2 := FALSE;
   B5_4.Word_buffer := 0;
   B5_4.Word_Result := 0;
   B5_5.Rising_Pulse_1 := FALSE;
   B5_5.Rising_Pulse_2 := FALSE;
   B5_5.Memory_Bit_1 := FALSE;
   B5_5.Memory_Bit_2 := FALSE;
   B5_5.Word_buffer := 0;
   B5_5.Word_Result := 0;
   B6_0.Rising_Pulse_1 := FALSE;
   B6_0.Rising_Pulse_2 := FALSE;
   B6_0.Memory_Bit_1 := FALSE;
   B6_0.Memory_Bit_2 := FALSE;
   B6_0.Word_buffer := 0;
   B6_0.Word_Result := 0;
   B6_1.Rising_Pulse_1 := FALSE;
   B6_1.Rising_Pulse_2 := FALSE;
   B6_1.Memory_Bit_1 := FALSE;
   B6_1.Memory_Bit_2 := FALSE;
   B6_1.Word_buffer := 0;
   B6_1.Word_Result := 0;
   B6_2.Rising_Pulse_1 := FALSE;
   B6_2.Rising_Pulse_2 := FALSE;
   B6_2.Memory_Bit_1 := FALSE;
   B6_2.Memory_Bit_2 := FALSE;
   B6_2.Word_buffer := 0;
   B6_2.Word_Result := 0;
   B6_4.Rising_Pulse_1 := FALSE;
   B6_4.Rising_Pulse_2 := FALSE;
   B6_4.Memory_Bit_1 := FALSE;
   B6_4.Memory_Bit_2 := FALSE;
   B6_4.Word_buffer := 0;
   B6_4.Word_Result := 0;
   B6_7.Rising_Pulse_1 := FALSE;
   B6_7.Rising_Pulse_2 := FALSE;
   B6_7.Memory_Bit_1 := FALSE;
   B6_7.Memory_Bit_2 := FALSE;
   B6_7.Word_buffer := 0;
   B6_7.Word_Result := 0;
   B7_0.Rising_Pulse_1 := FALSE;
   B7_0.Rising_Pulse_2 := FALSE;
   B7_0.Memory_Bit_1 := FALSE;
   B7_0.Memory_Bit_2 := FALSE;
   B7_0.Word_buffer := 0;
   B7_0.Word_Result := 0;
   B7_1.Rising_Pulse_1 := FALSE;
   B7_1.Rising_Pulse_2 := FALSE;
   B7_1.Memory_Bit_1 := FALSE;
   B7_1.Memory_Bit_2 := FALSE;
   B7_1.Word_buffer := 0;
   B7_1.Word_Result := 0;
   B7_2.Rising_Pulse_1 := FALSE;
   B7_2.Rising_Pulse_2 := FALSE;
   B7_2.Memory_Bit_1 := FALSE;
   B7_2.Memory_Bit_2 := FALSE;
   B7_2.Word_buffer := 0;
   B7_2.Word_Result := 0;
   B7_3.Rising_Pulse_1 := FALSE;
   B7_3.Rising_Pulse_2 := FALSE;
   B7_3.Memory_Bit_1 := FALSE;
   B7_3.Memory_Bit_2 := FALSE;
   B7_3.Word_buffer := 0;
   B7_3.Word_Result := 0;
   B7_4.Rising_Pulse_1 := FALSE;
   B7_4.Rising_Pulse_2 := FALSE;
   B7_4.Memory_Bit_1 := FALSE;
   B7_4.Memory_Bit_2 := FALSE;
   B7_4.Word_buffer := 0;
   B7_4.Word_Result := 0;
   B8_2.Rising_Pulse_1 := FALSE;
   B8_2.Rising_Pulse_2 := FALSE;
   B8_2.Memory_Bit_1 := FALSE;
   B8_2.Memory_Bit_2 := FALSE;
   B8_2.Word_buffer := 0;
   B8_2.Word_Result := 0;
   B9_6.Rising_Pulse_1 := FALSE;
   B9_6.Rising_Pulse_2 := FALSE;
   B9_6.Memory_Bit_1 := FALSE;
   B9_6.Memory_Bit_2 := FALSE;
   B9_6.Word_buffer := 0;
   B9_6.Word_Result := 0;
   B9_7.Rising_Pulse_1 := FALSE;
   B9_7.Rising_Pulse_2 := FALSE;
   B9_7.Memory_Bit_1 := FALSE;
   B9_7.Memory_Bit_2 := FALSE;
   B9_7.Word_buffer := 0;
   B9_7.Word_Result := 0;
   B10_3.Rising_Pulse_1 := FALSE;
   B10_3.Rising_Pulse_2 := FALSE;
   B10_3.Memory_Bit_1 := FALSE;
   B10_3.Memory_Bit_2 := FALSE;
   B10_3.Word_buffer := 0;
   B10_3.Word_Result := 0;
   B10_4.Rising_Pulse_1 := FALSE;
   B10_4.Rising_Pulse_2 := FALSE;
   B10_4.Memory_Bit_1 := FALSE;
   B10_4.Memory_Bit_2 := FALSE;
   B10_4.Word_buffer := 0;
   B10_4.Word_Result := 0;
   B10_5.Rising_Pulse_1 := FALSE;
   B10_5.Rising_Pulse_2 := FALSE;
   B10_5.Memory_Bit_1 := FALSE;
   B10_5.Memory_Bit_2 := FALSE;
   B10_5.Word_buffer := 0;
   B10_5.Word_Result := 0;
   B10_6.Rising_Pulse_1 := FALSE;
   B10_6.Rising_Pulse_2 := FALSE;
   B10_6.Memory_Bit_1 := FALSE;
   B10_6.Memory_Bit_2 := FALSE;
   B10_6.Word_buffer := 0;
   B10_6.Word_Result := 0;
   B10_7.Rising_Pulse_1 := FALSE;
   B10_7.Rising_Pulse_2 := FALSE;
   B10_7.Memory_Bit_1 := FALSE;
   B10_7.Memory_Bit_2 := FALSE;
   B10_7.Word_buffer := 0;
   B10_7.Word_Result := 0;
   B11_0.Rising_Pulse_1 := FALSE;
   B11_0.Rising_Pulse_2 := FALSE;
   B11_0.Memory_Bit_1 := FALSE;
   B11_0.Memory_Bit_2 := FALSE;
   B11_0.Word_buffer := 0;
   B11_0.Word_Result := 0;
   B11_1.Rising_Pulse_1 := FALSE;
   B11_1.Rising_Pulse_2 := FALSE;
   B11_1.Memory_Bit_1 := FALSE;
   B11_1.Memory_Bit_2 := FALSE;
   B11_1.Word_buffer := 0;
   B11_1.Word_Result := 0;
   B12_3.Rising_Pulse_1 := FALSE;
   B12_3.Rising_Pulse_2 := FALSE;
   B12_3.Memory_Bit_1 := FALSE;
   B12_3.Memory_Bit_2 := FALSE;
   B12_3.Word_buffer := 0;
   B12_3.Word_Result := 0;
   B13_0.Rising_Pulse_1 := FALSE;
   B13_0.Rising_Pulse_2 := FALSE;
   B13_0.Memory_Bit_1 := FALSE;
   B13_0.Memory_Bit_2 := FALSE;
   B13_0.Word_buffer := 0;
   B13_0.Word_Result := 0;
   B15_4.Rising_Pulse_1 := FALSE;
   B15_4.Rising_Pulse_2 := FALSE;
   B15_4.Memory_Bit_1 := FALSE;
   B15_4.Memory_Bit_2 := FALSE;
   B15_4.Word_buffer := 0;
   B15_4.Word_Result := 0;
   B15_5.Rising_Pulse_1 := FALSE;
   B15_5.Rising_Pulse_2 := FALSE;
   B15_5.Memory_Bit_1 := FALSE;
   B15_5.Memory_Bit_2 := FALSE;
   B15_5.Word_buffer := 0;
   B15_5.Word_Result := 0;
   B15_6.Rising_Pulse_1 := FALSE;
   B15_6.Rising_Pulse_2 := FALSE;
   B15_6.Memory_Bit_1 := FALSE;
   B15_6.Memory_Bit_2 := FALSE;
   B15_6.Word_buffer := 0;
   B15_6.Word_Result := 0;
   B15_7.Rising_Pulse_1 := FALSE;
   B15_7.Rising_Pulse_2 := FALSE;
   B15_7.Memory_Bit_1 := FALSE;
   B15_7.Memory_Bit_2 := FALSE;
   B15_7.Word_buffer := 0;
   B15_7.Word_Result := 0;
   B35_2.Rising_Pulse_1 := FALSE;
   B35_2.Rising_Pulse_2 := FALSE;
   B35_2.Memory_Bit_1 := FALSE;
   B35_2.Memory_Bit_2 := FALSE;
   B35_2.Word_buffer := 0;
   B35_2.Word_Result := 0;
   B35_3.Rising_Pulse_1 := FALSE;
   B35_3.Rising_Pulse_2 := FALSE;
   B35_3.Memory_Bit_1 := FALSE;
   B35_3.Memory_Bit_2 := FALSE;
   B35_3.Word_buffer := 0;
   B35_3.Word_Result := 0;
   B35_4.Rising_Pulse_1 := FALSE;
   B35_4.Rising_Pulse_2 := FALSE;
   B35_4.Memory_Bit_1 := FALSE;
   B35_4.Memory_Bit_2 := FALSE;
   B35_4.Word_buffer := 0;
   B35_4.Word_Result := 0;
   B11_2.Rising_Pulse_1 := FALSE;
   B11_2.Rising_Pulse_2 := FALSE;
   B11_2.Memory_Bit_1 := FALSE;
   B11_2.Memory_Bit_2 := FALSE;
   B11_2.Word_buffer := 0;
   B11_2.Word_Result := 0;
   Z2040 := FALSE;
   M052 := FALSE;
   M1122 := FALSE;
   M1123 := FALSE;
   M1124 := FALSE;
   M1125 := FALSE;
   M1126 := FALSE;
   M1127 := FALSE;
END_DATA_BLOCK

DATA_BLOCK "COLLATORS DB"
TITLE =
NAME : COLLATOR
VERSION : 0.1


  STRUCT
   SoftWare_Gate_0 : BOOL ;	//SoftWare Gate 0
   SoftWare_Gate_1 : BOOL ;	//SoftWare Gate 1
   SoftWare_Gate_2 : BOOL ;	//SoftWare Gate 2
   SoftWare_Gate_3 : BOOL ;	//SoftWare Gate 3
   SoftWare_Gate_4 : BOOL ;	//SoftWare Gate 4
   SoftWare_Gate_5 : BOOL ;	//SoftWare Gate 5
   SoftWare_Gate_6 : BOOL ;	//SoftWare Gate 6
   SoftWare_Gate_7 : BOOL ;	//SoftWare Gate 7
   DB_VAR8 : BOOL ;	//Temporary placeholder variable
   DB_VAR9 : BOOL ;	//Temporary placeholder variable
   DB_VAR10 : BOOL ;	//Temporary placeholder variable
   DB_VAR11 : BOOL ;	//Temporary placeholder variable
   DB_VAR12 : BOOL ;	//Temporary placeholder variable
   DB_VAR13 : BOOL ;	//Temporary placeholder variable
   DB_VAR14 : BOOL ;	//Temporary placeholder variable
   DB_VAR15 : BOOL ;	//Temporary placeholder variable
   Conveyor_Length_C3 : WORD ;	//Conveyor 3 - Conveyor Length (Fixed - Do Not Change !)
   Press_Length_C3 : WORD ;	//Conveyor 3 - Press Length
   DB_Conveyor_C3 : WORD ;	//Conveyor 3 - Spare
   DB_Conveyor_34 : WORD ;	//Conveyor 3 - Spare
   DB_Conveyor_31 : WORD ;	//Conveyor 3 - Spare
   Any_Conveyors_mS : DWORD ;	//Conveyor 3 - Any Conveyor mS TEST  [mS]
   DB_Conveyor_3321 : INT ;	//Conveyor 3 - Spare
   DB_Conveyor_33211 : INT ;	//Conveyor 3 - Spare
   Surface_Left_C4 : WORD ;	//Conveyor 4 - Surface_Left_Mem
   Frac_Packet_Length_C4 : WORD ;	//Conveyor 4 - Fraction of Packet Length
   PacketLength_C4 : WORD ;	//Conveyor 4 - Packet Length [Encoder Pulses]
   Packet_Length_Frac_C4 : WORD ;	//Conveyor 4 - Packet Length + Fraction [Encoder Pulses]
   Surface_Length_C4 : WORD ;	//Conveyor 4 - Surface Length [Encoder Pulses]
   Surface_Length_Left_C4 : WORD ;	//Conveyor 4 - Surface Length Remaining [Encoder Pulses]
   Spare_C4 : INT  := 635;	//Conveyor 4 - Spare
   Packet_Length_C4_mS : INT ;	//Conveyor 4 - Packet Length C4  [mS]
   Encoder_MM_Pulse_C4 : REAL ;	//Conveyor 4 - Encoder C4 [mm/pulse]
   Encoder_MM_Pulse_C10 : REAL ;	//Conveyor 10 - Encoder C10 [mm/pulse]
   DB_Conveyor_332121 : INT ;	//Conveyor 4 - Spare
   Frac_Packet_Width_C10 : WORD ;	//Conveyor 10 - Fraction of Packet Width [Encoder Pulses]
   Packet_Width_C10 : WORD ;	//Conveyor 10 - Packet Width [Encoder Pulses]
   Packet_Width_Frac_C10 : WORD ;	//Conveyor 10 - Packet Width + Fraction [Encoder Pulses]
   Surface_Length_10 : WORD ;	//Conveyor 10 - Surface Length [Encoder Pulses]
   Surface_Length_Left_10 : WORD ;	//Conveyor 10 - Surface Length Remaining [Encoder Pulses]
   Ecoder_Wheel_Circ_C10 : INT  := 283;	//Conveyor 10 - Encoder Wheel Circumference 283 mm
   Packet_Width_C10_mS : DWORD ;	//Conveyor 10 - Packet Width C10 [mS]
   DB_Conveyor_33232 : REAL ;	//Conveyor 10 - Spare
   DB_Conveyor_33233 : REAL ;	//Conveyor 10 - Spare
  END_STRUCT ;
BEGIN
   SoftWare_Gate_0 := FALSE;
   SoftWare_Gate_1 := FALSE;
   SoftWare_Gate_2 := FALSE;
   SoftWare_Gate_3 := FALSE;
   SoftWare_Gate_4 := FALSE;
   SoftWare_Gate_5 := FALSE;
   SoftWare_Gate_6 := FALSE;
   SoftWare_Gate_7 := FALSE;
   DB_VAR8 := FALSE;
   DB_VAR9 := FALSE;
   DB_VAR10 := FALSE;
   DB_VAR11 := FALSE;
   DB_VAR12 := FALSE;
   DB_VAR13 := FALSE;
   DB_VAR14 := FALSE;
   DB_VAR15 := FALSE;
   Conveyor_Length_C3 := W#16#0;
   Press_Length_C3 := W#16#0;
   DB_Conveyor_C3 := W#16#0;
   DB_Conveyor_34 := W#16#0;
   DB_Conveyor_31 := W#16#0;
   Any_Conveyors_mS := DW#16#0;
   DB_Conveyor_3321 := 0;
   DB_Conveyor_33211 := 0;
   Surface_Left_C4 := W#16#0;
   Frac_Packet_Length_C4 := W#16#0;
   PacketLength_C4 := W#16#0;
   Packet_Length_Frac_C4 := W#16#0;
   Surface_Length_C4 := W#16#0;
   Surface_Length_Left_C4 := W#16#0;
   Spare_C4 := 0;
   Packet_Length_C4_mS := 0;
   Encoder_MM_Pulse_C4 := 0.000000e+000;
   Encoder_MM_Pulse_C10 := 0.000000e+000;
   DB_Conveyor_332121 := 0;
   Frac_Packet_Width_C10 := W#16#0;
   Packet_Width_C10 := W#16#0;
   Packet_Width_Frac_C10 := W#16#0;
   Surface_Length_10 := W#16#0;
   Surface_Length_Left_10 := W#16#0;
   Ecoder_Wheel_Circ_C10 := 283;
   Packet_Width_C10_mS := DW#16#0;
   DB_Conveyor_33232 := 0.000000e+000;
   DB_Conveyor_33233 := 0.000000e+000;
END_DATA_BLOCK

DATA_BLOCK "DEBOUNCER COUNTER DB"
TITLE = DB8
VERSION : 0.1


  STRUCT
   Conveyor_C3_Slat : "Debouncer Counter Struct";	//C3 Struct
   Conveyor_C4_Collator : "Debouncer Counter Struct";	//C4 Struct
   Conveyor_C5_Link : "Debouncer Counter Struct";	//C5 Struct
   Conveyor_C6_Delivery : "Debouncer Counter Struct";	//C6 Struct
   Conveyor_C10_Collator : "Debouncer Counter Struct";	//C10 Struct
   Conveyor_C11_Link : "Debouncer Counter Struct";	//C11 Struct
   Conveyor_C12_Link : "Debouncer Counter Struct";	//C12 Struct
   Conveyor_C13_Delivery : "Debouncer Counter Struct";	//C13 Struct
   Conveyor_C21_Link : "Debouncer Counter Struct";	//C21 Struct
   Conveyor_C22_Link : "Debouncer Counter Struct";	//C22 Struct
   Conveyor_C23_Delivery : "Debouncer Counter Struct";	//C23 Struct
  END_STRUCT ;
BEGIN
   Conveyor_C3_Slat.FirstScan_Done := FALSE;
   Conveyor_C3_Slat.Bit0_ON_Latch := FALSE;
   Conveyor_C3_Slat.Bit1_ON_Latch := FALSE;
   Conveyor_C3_Slat.Transfer_Active := FALSE;
   Conveyor_C3_Slat.Count_Done_Latch_0 := FALSE;
   Conveyor_C3_Slat.Count_Done_Latch_1 := FALSE;
   Conveyor_C3_Slat.Error := FALSE;
   Conveyor_C3_Slat.Spare_Bit := FALSE;
   Conveyor_C3_Slat.Bit0_Entry_mS := 0;
   Conveyor_C3_Slat.Bit0_OFF_mS := 0;
   Conveyor_C3_Slat.Bit0_Stuck_mS := 0;
   Conveyor_C3_Slat.Bit1_Exit_mS := 0;
   Conveyor_C3_Slat.Bit1_OFF_mS := 0;
   Conveyor_C3_Slat.Space_Between := 0;
   Conveyor_C3_Slat.InFeed_Window_mS := 0;
   Conveyor_C3_Slat.Exit_Window_mS := 0;
   Conveyor_C3_Slat.Count_Result := 0;
   Conveyor_C3_Slat.Maximum_Count := 0;
   Conveyor_C3_Slat.HMI_Last := 0;
   Conveyor_C4_Collator.FirstScan_Done := FALSE;
   Conveyor_C4_Collator.Bit0_ON_Latch := FALSE;
   Conveyor_C4_Collator.Bit1_ON_Latch := FALSE;
   Conveyor_C4_Collator.Transfer_Active := FALSE;
   Conveyor_C4_Collator.Count_Done_Latch_0 := FALSE;
   Conveyor_C4_Collator.Count_Done_Latch_1 := FALSE;
   Conveyor_C4_Collator.Error := FALSE;
   Conveyor_C4_Collator.Spare_Bit := FALSE;
   Conveyor_C4_Collator.Bit0_Entry_mS := 0;
   Conveyor_C4_Collator.Bit0_OFF_mS := 0;
   Conveyor_C4_Collator.Bit0_Stuck_mS := 0;
   Conveyor_C4_Collator.Bit1_Exit_mS := 0;
   Conveyor_C4_Collator.Bit1_OFF_mS := 0;
   Conveyor_C4_Collator.Space_Between := 0;
   Conveyor_C4_Collator.InFeed_Window_mS := 0;
   Conveyor_C4_Collator.Exit_Window_mS := 0;
   Conveyor_C4_Collator.Count_Result := 0;
   Conveyor_C4_Collator.Maximum_Count := 0;
   Conveyor_C4_Collator.HMI_Last := 0;
   Conveyor_C5_Link.FirstScan_Done := FALSE;
   Conveyor_C5_Link.Bit0_ON_Latch := FALSE;
   Conveyor_C5_Link.Bit1_ON_Latch := FALSE;
   Conveyor_C5_Link.Transfer_Active := FALSE;
   Conveyor_C5_Link.Count_Done_Latch_0 := FALSE;
   Conveyor_C5_Link.Count_Done_Latch_1 := FALSE;
   Conveyor_C5_Link.Error := FALSE;
   Conveyor_C5_Link.Spare_Bit := FALSE;
   Conveyor_C5_Link.Bit0_Entry_mS := 0;
   Conveyor_C5_Link.Bit0_OFF_mS := 0;
   Conveyor_C5_Link.Bit0_Stuck_mS := 0;
   Conveyor_C5_Link.Bit1_Exit_mS := 0;
   Conveyor_C5_Link.Bit1_OFF_mS := 0;
   Conveyor_C5_Link.Space_Between := 0;
   Conveyor_C5_Link.InFeed_Window_mS := 0;
   Conveyor_C5_Link.Exit_Window_mS := 0;
   Conveyor_C5_Link.Count_Result := 0;
   Conveyor_C5_Link.Maximum_Count := 0;
   Conveyor_C5_Link.HMI_Last := 0;
   Conveyor_C6_Delivery.FirstScan_Done := FALSE;
   Conveyor_C6_Delivery.Bit0_ON_Latch := FALSE;
   Conveyor_C6_Delivery.Bit1_ON_Latch := FALSE;
   Conveyor_C6_Delivery.Transfer_Active := FALSE;
   Conveyor_C6_Delivery.Count_Done_Latch_0 := FALSE;
   Conveyor_C6_Delivery.Count_Done_Latch_1 := FALSE;
   Conveyor_C6_Delivery.Error := FALSE;
   Conveyor_C6_Delivery.Spare_Bit := FALSE;
   Conveyor_C6_Delivery.Bit0_Entry_mS := 0;
   Conveyor_C6_Delivery.Bit0_OFF_mS := 0;
   Conveyor_C6_Delivery.Bit0_Stuck_mS := 0;
   Conveyor_C6_Delivery.Bit1_Exit_mS := 0;
   Conveyor_C6_Delivery.Bit1_OFF_mS := 0;
   Conveyor_C6_Delivery.Space_Between := 0;
   Conveyor_C6_Delivery.InFeed_Window_mS := 0;
   Conveyor_C6_Delivery.Exit_Window_mS := 0;
   Conveyor_C6_Delivery.Count_Result := 0;
   Conveyor_C6_Delivery.Maximum_Count := 0;
   Conveyor_C6_Delivery.HMI_Last := 0;
   Conveyor_C10_Collator.FirstScan_Done := FALSE;
   Conveyor_C10_Collator.Bit0_ON_Latch := FALSE;
   Conveyor_C10_Collator.Bit1_ON_Latch := FALSE;
   Conveyor_C10_Collator.Transfer_Active := FALSE;
   Conveyor_C10_Collator.Count_Done_Latch_0 := FALSE;
   Conveyor_C10_Collator.Count_Done_Latch_1 := FALSE;
   Conveyor_C10_Collator.Error := FALSE;
   Conveyor_C10_Collator.Spare_Bit := FALSE;
   Conveyor_C10_Collator.Bit0_Entry_mS := 0;
   Conveyor_C10_Collator.Bit0_OFF_mS := 0;
   Conveyor_C10_Collator.Bit0_Stuck_mS := 0;
   Conveyor_C10_Collator.Bit1_Exit_mS := 0;
   Conveyor_C10_Collator.Bit1_OFF_mS := 0;
   Conveyor_C10_Collator.Space_Between := 0;
   Conveyor_C10_Collator.InFeed_Window_mS := 0;
   Conveyor_C10_Collator.Exit_Window_mS := 0;
   Conveyor_C10_Collator.Count_Result := 0;
   Conveyor_C10_Collator.Maximum_Count := 0;
   Conveyor_C10_Collator.HMI_Last := 0;
   Conveyor_C11_Link.FirstScan_Done := FALSE;
   Conveyor_C11_Link.Bit0_ON_Latch := FALSE;
   Conveyor_C11_Link.Bit1_ON_Latch := FALSE;
   Conveyor_C11_Link.Transfer_Active := FALSE;
   Conveyor_C11_Link.Count_Done_Latch_0 := FALSE;
   Conveyor_C11_Link.Count_Done_Latch_1 := FALSE;
   Conveyor_C11_Link.Error := FALSE;
   Conveyor_C11_Link.Spare_Bit := FALSE;
   Conveyor_C11_Link.Bit0_Entry_mS := 0;
   Conveyor_C11_Link.Bit0_OFF_mS := 0;
   Conveyor_C11_Link.Bit0_Stuck_mS := 0;
   Conveyor_C11_Link.Bit1_Exit_mS := 0;
   Conveyor_C11_Link.Bit1_OFF_mS := 0;
   Conveyor_C11_Link.Space_Between := 0;
   Conveyor_C11_Link.InFeed_Window_mS := 0;
   Conveyor_C11_Link.Exit_Window_mS := 0;
   Conveyor_C11_Link.Count_Result := 0;
   Conveyor_C11_Link.Maximum_Count := 0;
   Conveyor_C11_Link.HMI_Last := 0;
   Conveyor_C12_Link.FirstScan_Done := FALSE;
   Conveyor_C12_Link.Bit0_ON_Latch := FALSE;
   Conveyor_C12_Link.Bit1_ON_Latch := FALSE;
   Conveyor_C12_Link.Transfer_Active := FALSE;
   Conveyor_C12_Link.Count_Done_Latch_0 := FALSE;
   Conveyor_C12_Link.Count_Done_Latch_1 := FALSE;
   Conveyor_C12_Link.Error := FALSE;
   Conveyor_C12_Link.Spare_Bit := FALSE;
   Conveyor_C12_Link.Bit0_Entry_mS := 0;
   Conveyor_C12_Link.Bit0_OFF_mS := 0;
   Conveyor_C12_Link.Bit0_Stuck_mS := 0;
   Conveyor_C12_Link.Bit1_Exit_mS := 0;
   Conveyor_C12_Link.Bit1_OFF_mS := 0;
   Conveyor_C12_Link.Space_Between := 0;
   Conveyor_C12_Link.InFeed_Window_mS := 0;
   Conveyor_C12_Link.Exit_Window_mS := 0;
   Conveyor_C12_Link.Count_Result := 0;
   Conveyor_C12_Link.Maximum_Count := 0;
   Conveyor_C12_Link.HMI_Last := 0;
   Conveyor_C13_Delivery.FirstScan_Done := FALSE;
   Conveyor_C13_Delivery.Bit0_ON_Latch := FALSE;
   Conveyor_C13_Delivery.Bit1_ON_Latch := FALSE;
   Conveyor_C13_Delivery.Transfer_Active := FALSE;
   Conveyor_C13_Delivery.Count_Done_Latch_0 := FALSE;
   Conveyor_C13_Delivery.Count_Done_Latch_1 := FALSE;
   Conveyor_C13_Delivery.Error := FALSE;
   Conveyor_C13_Delivery.Spare_Bit := FALSE;
   Conveyor_C13_Delivery.Bit0_Entry_mS := 0;
   Conveyor_C13_Delivery.Bit0_OFF_mS := 0;
   Conveyor_C13_Delivery.Bit0_Stuck_mS := 0;
   Conveyor_C13_Delivery.Bit1_Exit_mS := 0;
   Conveyor_C13_Delivery.Bit1_OFF_mS := 0;
   Conveyor_C13_Delivery.Space_Between := 0;
   Conveyor_C13_Delivery.InFeed_Window_mS := 0;
   Conveyor_C13_Delivery.Exit_Window_mS := 0;
   Conveyor_C13_Delivery.Count_Result := 0;
   Conveyor_C13_Delivery.Maximum_Count := 0;
   Conveyor_C13_Delivery.HMI_Last := 0;
   Conveyor_C21_Link.FirstScan_Done := FALSE;
   Conveyor_C21_Link.Bit0_ON_Latch := FALSE;
   Conveyor_C21_Link.Bit1_ON_Latch := FALSE;
   Conveyor_C21_Link.Transfer_Active := FALSE;
   Conveyor_C21_Link.Count_Done_Latch_0 := FALSE;
   Conveyor_C21_Link.Count_Done_Latch_1 := FALSE;
   Conveyor_C21_Link.Error := FALSE;
   Conveyor_C21_Link.Spare_Bit := FALSE;
   Conveyor_C21_Link.Bit0_Entry_mS := 0;
   Conveyor_C21_Link.Bit0_OFF_mS := 0;
   Conveyor_C21_Link.Bit0_Stuck_mS := 0;
   Conveyor_C21_Link.Bit1_Exit_mS := 0;
   Conveyor_C21_Link.Bit1_OFF_mS := 0;
   Conveyor_C21_Link.Space_Between := 0;
   Conveyor_C21_Link.InFeed_Window_mS := 0;
   Conveyor_C21_Link.Exit_Window_mS := 0;
   Conveyor_C21_Link.Count_Result := 0;
   Conveyor_C21_Link.Maximum_Count := 0;
   Conveyor_C21_Link.HMI_Last := 0;
   Conveyor_C22_Link.FirstScan_Done := FALSE;
   Conveyor_C22_Link.Bit0_ON_Latch := FALSE;
   Conveyor_C22_Link.Bit1_ON_Latch := FALSE;
   Conveyor_C22_Link.Transfer_Active := FALSE;
   Conveyor_C22_Link.Count_Done_Latch_0 := FALSE;
   Conveyor_C22_Link.Count_Done_Latch_1 := FALSE;
   Conveyor_C22_Link.Error := FALSE;
   Conveyor_C22_Link.Spare_Bit := FALSE;
   Conveyor_C22_Link.Bit0_Entry_mS := 0;
   Conveyor_C22_Link.Bit0_OFF_mS := 0;
   Conveyor_C22_Link.Bit0_Stuck_mS := 0;
   Conveyor_C22_Link.Bit1_Exit_mS := 0;
   Conveyor_C22_Link.Bit1_OFF_mS := 0;
   Conveyor_C22_Link.Space_Between := 0;
   Conveyor_C22_Link.InFeed_Window_mS := 0;
   Conveyor_C22_Link.Exit_Window_mS := 0;
   Conveyor_C22_Link.Count_Result := 0;
   Conveyor_C22_Link.Maximum_Count := 0;
   Conveyor_C22_Link.HMI_Last := 0;
   Conveyor_C23_Delivery.FirstScan_Done := FALSE;
   Conveyor_C23_Delivery.Bit0_ON_Latch := FALSE;
   Conveyor_C23_Delivery.Bit1_ON_Latch := FALSE;
   Conveyor_C23_Delivery.Transfer_Active := FALSE;
   Conveyor_C23_Delivery.Count_Done_Latch_0 := FALSE;
   Conveyor_C23_Delivery.Count_Done_Latch_1 := FALSE;
   Conveyor_C23_Delivery.Error := FALSE;
   Conveyor_C23_Delivery.Spare_Bit := FALSE;
   Conveyor_C23_Delivery.Bit0_Entry_mS := 0;
   Conveyor_C23_Delivery.Bit0_OFF_mS := 0;
   Conveyor_C23_Delivery.Bit0_Stuck_mS := 0;
   Conveyor_C23_Delivery.Bit1_Exit_mS := 0;
   Conveyor_C23_Delivery.Bit1_OFF_mS := 0;
   Conveyor_C23_Delivery.Space_Between := 0;
   Conveyor_C23_Delivery.InFeed_Window_mS := 0;
   Conveyor_C23_Delivery.Exit_Window_mS := 0;
   Conveyor_C23_Delivery.Count_Result := 0;
   Conveyor_C23_Delivery.Maximum_Count := 0;
   Conveyor_C23_Delivery.HMI_Last := 0;
END_DATA_BLOCK

DATA_BLOCK "HOUSE_KEEPING DB"
TITLE =
VERSION : 0.1


  STRUCT
   C4_First_Collating : BOOL ;	//C4 First Packet Collating
   C4_First_Collating_Done : BOOL ;	//C4 First Packet Collating Done
   C10_First_Collating : BOOL ;	//C10 First Packet Collating
   C10_First_Collating_Done : BOOL ;	//C10 First Packet Collating Done
   Spare5 : BOOL ;
   Spare6 : BOOL ;
   Spare7 : BOOL ;
   Spare8 : BOOL ;
   SpareWord : WORD ;
   C4_Added_Scans_mS : INT ;	//C4 Added Scan Cycles [mS]
   C10_Added_Scans_mS : INT ;	//C10 Added Scan Cycles [mS]
   C3_Encoder_READ_Mem : INT ;	//C3 Encoder Read / Print [ep](Encoder Pulses)
   C4_Encoder_READ_Mem : INT ;	//C4 Encoder Read / Print [ep](Encoder Pulses)
   C10_Encoder_READ_Mem : INT ;	//C10 Encoder Read / Print [ep](Encoder Pulses)
   C3_Packet_Length_ep : INT ;	//C3 Encoder Length [ep]
   C4_Packet_Length_ep : INT ;	//C4 Encoder Length [ep]
   C10_Packet_Width_ep : INT ;	//C10 Encoder Length [ep]
   C3_Packet_Length_mm : INT ;	//C3 Packet Lenght [mm]
   C4_Packet_Length_mm : INT ;	//C4 Packet Lenght [mm]
   C10_Packet_Width_mm : INT ;	//C10 Packet Lenght [mm]
   C4_Packet_Length_mS : INT ;	//C4 Packet Lenght [mS]
   C10_Packet_Width_mS : INT ;	//C4 Packet Lenght [mS]
   C4_RampDown_Dx_ep : INT ;	//C4 Ramp Down Distance [EP]
   C10_RampDown_Dx_ep : INT ;	//C10 Ramp Up/Down Distance [EP]
   SpareINT01 : INT ;
   SpareINT02 : INT ;
   SpareINT03 : INT ;
   SpareINT04 : INT ;
  END_STRUCT ;
BEGIN
   C4_First_Collating := FALSE;
   C4_First_Collating_Done := FALSE;
   C10_First_Collating := FALSE;
   C10_First_Collating_Done := FALSE;
   Spare5 := FALSE;
   Spare6 := FALSE;
   Spare7 := FALSE;
   Spare8 := FALSE;
   SpareWord := W#16#0;
   C4_Added_Scans_mS := 0;
   C10_Added_Scans_mS := 0;
   C3_Encoder_READ_Mem := 0;
   C4_Encoder_READ_Mem := 0;
   C10_Encoder_READ_Mem := 0;
   C3_Packet_Length_ep := 0;
   C4_Packet_Length_ep := 0;
   C10_Packet_Width_ep := 0;
   C3_Packet_Length_mm := 0;
   C4_Packet_Length_mm := 654;
   C10_Packet_Width_mm := 0;
   C4_Packet_Length_mS := 0;
   C10_Packet_Width_mS := 0;
   C4_RampDown_Dx_ep := 0;
   C10_RampDown_Dx_ep := 0;
   SpareINT01 := 0;
   SpareINT02 := 0;
   SpareINT03 := 0;
   SpareINT04 := 0;
END_DATA_BLOCK

DATA_BLOCK "HMI_DB"
TITLE =
VERSION : 0.1


  STRUCT
   GRAPHIC_INIT : BOOL ;	//FL Graphic Init
   EMERGENCY_BLINK : BOOL ;	//FL Emergency Blink
   TRANS_SYSTEM_ON_SW : BOOL ;	//FLS On Sw Temporary
   COMPRESSED_AIR : BOOL ;	//FLS Compressed Air
   TRANS_SYSTEM_RUN_STATUS : BOOL ;	//FLS 508 Link Run SW - Diabled
   PACKET_in_FLIPPER_SW : BOOL ;	//FLS Service Enable Switch - Disabled
   SERVICE_INIT_PB : BOOL ;	//FLS Service Initialisation PB
   ALL_SERVICE_ENABLE_SW : BOOL ;	//FLS All Services Enable Switch
   SERVICE_SW_1_STATUS : BOOL ;	//FLS Service 1 Switch
   SERVICE_SW_2_STATUS : BOOL ;	//FLS Service 2 Switch
   SERVICE_SW_3_STATUS : BOOL ;	//FLS Service 3 Switch
   SERVICE_SW_1_2_STATUS : BOOL ;	//FLS Service 1 or 2 Switch
   BIT12 : BOOL ;	//FLS Spare
   BIT13 : BOOL ;	//FLS Spare
   SERVICE_SW_2_TIME_ADJ : BOOL ;	//FLS Service 2 Switch - Time Adjust
   PACKETIZER_GATE_STATUS : BOOL ;	//FLS 2145 Packetizer Flap Gate - Status Bit
   E_STOP_CONSOLE_STATUS : BOOL ;	//FL E-Stop Console
   E_STOP_ELEVATOR_STATUS : BOOL ;	//FL E-Stop Elevator
   E_STOP_FLIPPER_STATUS : BOOL ;	//FL E-Stop Flipper
   E_STOP_LOADER_STATUS : BOOL ;	//FL E-Stop Loader
   HAND_FEED_ARROW_STATUS : BOOL ;	//FL Hand Feed Arrow
   ELEVATOR_DOOR_STATUS : BOOL ;	//FL Elevator Door
   FLIPPER_DOOR_STATUS : BOOL ;	//FL Flipper Door
   LOADER_DOOR_STATUS : BOOL ;	//FL Loader Door
   LIGHT_BARRIER_1_STATUS : BOOL ;	//FL Light Barrier 1 - B5.4 Conveyor 1 Exit - Status Bit
   LIGHT_BARRIER_2_STATUS : BOOL ;	//FL Light Barrier 2 - B5.5 Conveyor 2 InFeed - Status Bit
   LIGHT_BARRIER_3_STATUS : BOOL ;	//FL Light Barrier 3 - B6.0 Conveyor 2 Presence - Status Bit
   LIGHT_BARRIER_4_STATUS : BOOL ;	//FL Light Barrier 4 - B6.1 Conveyor 2 Exit - Status Bit
   LIGHT_BARRIER_5_STATUS : BOOL ;	//FL Light Barrier 5 - B6.2 Conveyor 3 InFeed - Status Bit
   LIGHT_BARRIER_6_STATUS : BOOL ;	//FL Light Barrier 6 - B6.4 Conveyor 3 Exit - Status Bit
   LIGHT_BARRIER_B_STATUS : BOOL ;	//FL Light Barrier B - B5.2 Elevator Limit - Status Bit
   LIGHT_BARRIER_A_STATUS : BOOL ;	//FL Light Barrier A - B5.1 Elevator InFeed - Status Bit
   BIT32 : BOOL ;	//FL Pusher 0 Motion
   BIT33 : BOOL ;	//FL Pusher 0 Motion
   BIT34 : BOOL ;	//FL Pusher 0 Motion
   BIT35 : BOOL ;	//FL Pusher 0 Motion
   BIT36 : BOOL ;	//FL Pusher 0 Motion
   BIT37 : BOOL ;	//FL Pusher 0 Motion
   BIT38 : BOOL ;	//FL Pusher 0 Motion
   BIT39 : BOOL ;	//FL Pusher 0 Motion
   BIT40 : BOOL ;	//FL Elevator Motion
   BIT41 : BOOL ;	//FL Elevator Motion
   BIT42 : BOOL ;	//FL Elevator Motion
   BIT43 : BOOL ;	//FL Elevator Motion
   BIT44 : BOOL ;	//FL Elevator Motion
   BIT45 : BOOL ;	//FL Elevator Motion
   BIT46 : BOOL ;	//FL Elevator Motion
   BIT47 : BOOL ;	//FL Elevator Motion
   BIT48 : BOOL ;	//FL Pusher 1 Motion
   BIT49 : BOOL ;	//FL Pusher 1 Motion
   BIT50 : BOOL ;	//FL Pusher 1 Motion
   BIT51 : BOOL ;	//FL Pusher 1 Motion
   BIT52 : BOOL ;	//FL Pusher 1 Motion
   BIT53 : BOOL ;	//FL Pusher 1 Motion
   BIT54 : BOOL ;	//FL Pusher 1 Motion
   BIT55 : BOOL ;	//FL Pusher 1 Motion
   BIT56 : BOOL ;	//FL Pusher 2 Motion
   BIT57 : BOOL ;	//FL Pusher 2 Motion
   BIT58 : BOOL ;	//FL Pusher 2 Motion
   BIT59 : BOOL ;	//FL Pusher 2 Motion
   BIT60 : BOOL ;	//FL Pusher 2 Motion
   BIT61 : BOOL ;	//FL Pusher 2 Motion
   BIT62 : BOOL ;	//FL Pusher 2 Motion
   CONVEYORS_CLEARING : BOOL ;	//FL Conveyors Clearing
   ELEVATOR_MOTOR_STATUS : BOOL ;	//FL Elevator - Motor M42.0 Status Bit
   PUSHER_1_MOTOR_STATUS : BOOL ;	//FL Pusher 1 - Motor M42.6 Status Bit
   CONVEYOR_1_MOTOR_STATUS : BOOL ;	//FL Conv 1 - Motor M43.0 Status Bit
   CONVEYOR_2B_MOTOR_STATUS : BOOL ;	//FL Conv 2 Belt - Motor M43.4 Status Bit
   CONVEYOR_2R_MOTOR_STATUS : BOOL ;	//FL Conv 2 Roller - Motor M43.5 Status Bit
   CONVEYOR_3_MOTOR_STATUS : BOOL ;	//FL Conveyor 3 - Motor M44.0 Status Bit
   CONVEYOR_4_MOTOR_STATUS : BOOL ;	//FL Conveyor 4 - Motor M44.3 Status Bit
   CONVEYOR_5_MOTOR_STATUS : BOOL ;	//FL Conveyor 5 - Motor M45.0 Status Bit
   CONVEYOR_6_MOTOR_STATUS : BOOL ;	//FL Conveyor 6 - Motor M45.3 Status Bit
   CONVEYOR_7_MOTOR_STATUS : BOOL ;	//FL Conveyor 7 - Motor M45.6 Status Bit
   FLIPPER_MOTOR_STATUS : BOOL ;	//FL Flipper Flip - Motor M46.0 Status Bit
   CONVEYOR_8_MOTOR_STATUS : BOOL ;	//FL Conveyor 8 - Motor M46.4 Status Bit
   TURNTABLE_MOTOR_STATUS : BOOL ;	//FL TurnTable - Motor M47.0 Status Bit
   CONVEYOR_9_MOTOR_STATUS : BOOL ;	//FL Conveyor 9 - Motor M47.5 Status Bit
   PUSHER_2_MOTOR_STATUS : BOOL ;	//FL Pusher 2 - Motor M47.6 Status Bit
   CONVEYOR_10_MOTOR_STATUS : BOOL ;	//FL Conveyor 10 - Motor M48.0 Status Bit
   CONVEYOR_11_MOTOR_STATUS : BOOL ;	//FL Conveyor 11 - Motor M48.3 Status Bit
   CONVEYOR_12_MOTOR_STATUS : BOOL ;	//FL Conveyor 12 - Motor M48.6 Status Bit
   CONVEYOR_13_MOTOR_STATUS : BOOL ;	//FL Conveyor 13 - Motor M49.0 Status Bit
   CONVEYOR_21_MOTOR_STATUS : BOOL ;	//FL Conveyor 21 - Motor M53.2 Status Bit
   CONVEYOR_22_MOTOR_STATUS : BOOL ;	//FL Conveyor 22 - Motor M53.4 Status Bit
   CONVEYOR_23_MOTOR_STATUS : BOOL ;	//FL Conveyor 23 - Motor M54.0 Status Bit
   LOADER_LIFT_MOTOR_STATUS : BOOL ;	//FL Loader Lift - Motor M50.0 Status Bit
   LOADER_FING_MOTOR_STATUS : BOOL ;	//FL Loader Fingers - Motor M50.5 Status Bit
   LOADER_BELT_MOTOR_STATUS : BOOL ;	//FL Loader Belt - Motor M51.0 Status Bit
   LIGHT_BARRIER_7_STATUS : BOOL ;	//FL Light Barrier 7 - B6.7 Conv 4 InFeed Sens - Status
   LIGHT_BARRIER_8_STATUS : BOOL ;	//FL Light Barrier 8 - B7.0 Conv 4 Exit Sens - Status
   LIGHT_BARRIER_9_STATUS : BOOL ;	//FL Light Barrier 9 - B7.1 Conv 5 Exit Sens - Status
   LIGHT_BARRIER_10_STATUS : BOOL ;	//FL Light Barrier 10 - B7.2 Conv 6 Slow Sens - Status Bit
   LIGHT_BARRIER_11_STATUS : BOOL ;	//FL Light Barrier 11 - B7.3 Conv 6 Exit Sens - Status Bit
   LIGHT_BARRIER_12_STATUS : BOOL ;	//FL Light Barrier 12 - B7.4 Flipper InFeed Sens - Status Bit
   LIGHT_BARRIER_13_STATUS : BOOL ;	//FL Light Barrier 13 - B8.2 Flipper Exit Sens - Status Bit
   LIGHT_BARRIER_14_STATUS : BOOL ;	//FL Light Barrier 14 - B9.6 Conv 9 InFeed Sens - Status Bit
   LIGHT_BARRIER_15_STATUS : BOOL ;	//FL Light Barrier 15 - B9.7 Conv 9 Packet Sens - Status Bit
   LIGHT_BARRIER_16_STATUS : BOOL ;	//FL Light Barrier 16 - B10.3 Conv 10 Start Sens - Status Bit
   LIGHT_BARRIER_17_STATUS : BOOL ;	//FL Light Barrier 17 - B10.4 Conv 10 InFeed Sens - Status Bit
   LIGHT_BARRIER_18_STATUS : BOOL ;	//FL Light Barrier 18 - B10.5 Conv 10 Full Sens - Status Bit
   LIGHT_BARRIER_19_STATUS : BOOL ;	//FL Light Barrier 19 - B10.6 Conv 10 Exit Sens - Status Bit
   LIGHT_BARRIER_20_STATUS : BOOL ;	//FL Light Barrier 20 - B10.7 Conv 11 Exit Sens - Status Bit
   LIGHT_BARRIER_21_STATUS : BOOL ;	//FL Light Barrier 21 - B11.0 Conv 12 Exit Sens - Status Bit- Status Bit
   LIGHT_BARRIER_22_STATUS : BOOL ;	//FL Light Barrier 22 - B11.1 Conv 13 Slow Sens - Status Bit
   LIGHT_BARRIER_23_STATUS : BOOL ;	//FL Light Barrier 23 - B11.2 Conv 13 Exit Sens - Status Bit
   LIGHT_BARRIER_24_STATUS : BOOL ;	//FL Light Barrier 24 - B12.3 Fingers Delivery Sens - Status Bit
   LIGHT_BARRIER_25_STATUS : BOOL ;	//FL Light Barrier 25 - B13.0 Loader Empty Sens - Status Bit
   LIGHT_BARRIER_26_STATUS : BOOL ;	//FL Light Barrier 26 - B15.4 Conv 21 Exit Sens - Status Bit
   LIGHT_BARRIER_27_STATUS : BOOL ;	//FL Light Barrier 27 - B15.5 Conv 22 Exit Sens - Status Bit
   LIGHT_BARRIER_28_STATUS : BOOL ;	//FL Light Barrier 28 - B15.6 Conv 23 Slow Sens - Status Bit
   LIGHT_BARRIER_29_STATUS : BOOL ;	//FL Light Barrier 29 - B15.7 Conv 23 Exit Sens - Status Bit
   LIGHT_BARRIER_30_STATUS : BOOL ;	//FL Light Barrier 30 - B35.2 Conv 0 InFeed Sens - Status Bit
   LIGHT_BARRIER_31_STATUS : BOOL ;	//FL Light Barrier 31 - B35.3 Conv 0 Exit Sens - Status Bit
   LIGHT_BARRIER_32_STATUS : BOOL ;	//FL Light Barrier 32 - B35.4 Conv 0 Length Sens - Status Bit
   PROX_9_STATUS : BOOL ;	//FL Prox 9 - P8.5 TurnTable Rotation InFeed Slow - Status Bit
   PROX_10_STATUS : BOOL ;	//FL Prox 10 - P8.6 TurnTable Rotation InFeed Stop - Status Bit
   PROX_11_STATUS : BOOL ;	//FL Prox 11 - P9.2 TurnTable Rotation Exit Slow - Status Bit
   PROX_12_STATUS : BOOL ;	//FL Prox 12 - P9.3 TurnTable Rotation Exit Stop - Status Bit
   PROX_13_STATUS : BOOL ;	//FL Prox 13 - P10.0 Pusher 2 Retract Sens - Status Bit
   PROX_14_STATUS : BOOL ;	//FL Prox 14 - P10.1 Pusher 2 Extend Sens - Status Bit
   PROX_15_STATUS : BOOL ;	//FL Prox 15 - P15.0 Pivot 10 High Sens - Status Bit
   PROX_16_STATUS : BOOL ;	//FL Prox 16 - P15.1 Pivot 10 Low Sens - Status Bit
   PROX_17_STATUS : BOOL ;	//FL Prox 17 - P13.2 Loader H Level Stop - Status Bit
   PROX_18_STATUS : BOOL ;	//FL Prox 18 - P13.1 Loader H Level Slow - Status Bit
   PROX_19_STATUS : BOOL ;	//FL Prox 19 - P11.4 Loader L Level Stop - Status Bit
   PROX_20_STATUS : BOOL ;	//FL Prox 20 - P11.5 Loader L Level Slow - Status Bit
   PROX_21_STATUS : BOOL ;	//FL Prox 21 - P11.6 Loader Slow Bot - Status Bit
   PROX_22_STATUS : BOOL ;	//FL Prox 22 - P11.7 Loader Stop Bot - Status Bit
   PROX_23_STATUS : BOOL ;	//FL Prox 23 - P12.0 Loader Finger Retract - Status Bit
   PROX_24_STATUS : BOOL ;	//FL Prox 24 - P12.1 Loader Finger Extend - Status Bit
   FP131 : BOOL ;	//FP One Shot
   FP132 : BOOL ;	//FP One Shot
   FP133 : BOOL ;	//FP One Shot
   FP134 : BOOL ;	//FP One Shot
   FP135 : BOOL ;	//FP One Shot
   TURNTABLE_DELIV_POSITION : BOOL ;	//FL TurnTable Delivery Position
   TURNTABLE_REVERSE_ARROW : BOOL ;	//FL TurnTable Arrow Reverse Packet
   TURNTABLE_DIR_SELECT_SW : BOOL ;	//FL TurnTable Direction Select SW
   TURNTABLE_FLICK_MOTION : BOOL ;	//FL TurnTable Flicker - Motion
   FP140 : BOOL ;	//FP One Shot
   FP141 : BOOL ;	//FP One Shot
   FP142 : BOOL ;	//FP One Shot
   FP143 : BOOL ;	//FP One Shot
   PROX_1_STATUS : BOOL ;	//FL Prox 1 - P4.0 Elevator Bottom Position - Status Bit
   PROX_2_STATUS : BOOL ;	//FL Prox 2 - P4.1 Elevator SlowDown Bot - Status Bit
   PROX_3_STATUS : BOOL ;	//FL Prox 3 - P4.2 Elevator SlowDown Top - Status Bit
   PROX_4_STATUS : BOOL ;	//FL Prox 4 - P4.3 Elevator Top Position - Status Bit
   PROX_5_STATUS : BOOL ;	//FL Prox 5 - P4.4 Pusher 1 Home - Status Bit
   PROX_6_STATUS : BOOL ;	//FL Prox 6 - P4.5 Pusher 1 Limit - Status Bit
   PROX_7_STATUS : BOOL ;	//FL Prox 7 - P8.0 Flipper Fingers Right Position - Status Bit
   PROX_8_STATUS : BOOL ;	//FL Prox 8 - P8.1 Flipper Fingers Left Position - Status Bit
   BIT152 : BOOL ;	//FL Loader Motion
   BIT153 : BOOL ;	//FL Loader Motion
   BIT154 : BOOL ;	//FL Loader Motion
   BIT155 : BOOL ;	//FL Loader Motion
   BIT156 : BOOL ;	//FL Loader Motion
   BIT157 : BOOL ;	//FL Loader Motion
   BIT158 : BOOL ;	//FL Loader Motion
   BIT159 : BOOL ;	//FL Loader Motion
   SERVICE_SSW_MAIN : BOOL ;	//FL Service SW Main Screen
   SERVICE_SSW_STATUS : BOOL ;	//FL Service SW Main Screen - Status
   CLEARING_SSW_MAIN : BOOL ;	//FL Clearing SW Main Screen
   CLEARING_SSW_STATUS : BOOL ;	//FL Clearing SW Main Screen - Status
   MAN_FEED_SSW_MAIN : BOOL ;	//FL Hand Feed SW Main Screen
   MAN_FEED_SSW_STATUS : BOOL ;	//FL Hand Feed SW Main Screen - Status
   TURNTABLE_SSW_MAIN : BOOL ;	//FL Turn Table Turn SW = 1:CCW - 0:CW Main Screen
   TURNTABLE_SSW_STATUS : BOOL ;	//FL Turn Table Select Main Screen - Status
   FLIPPER_SSW_MAIN : BOOL ;	//FL Flipper SW Main Screen
   FLIPPER_SSW_STATUS : BOOL ;	//FL Flipper SW Main Screen - Status
   ROLLER_SSW_MAIN : BOOL ;	//FL Roller SW Main Screen
   ROLLER_SSW_STATUS : BOOL ;	//FL Roller SW Main Screen - Status
   ELEVATOR_ROUND_TRIP_SSW : BOOL ;	//FL Elevator - Round Trip PB
   BIT173 : BOOL ;
   BIT174 : BOOL ;
   BIT175 : BOOL ;
   HMI_PUSHER_0_TEST_SSW : BOOL ;	//FL Pusher 0 SW
   HMI_ELEVATOR_SERVICE_SSW : BOOL ;	//FL Elevator Service SW
   HMI_ELEVATOR_TEST_DN_SSW : BOOL ;	//FL Elevator DN PB
   HMI_ELEVATOR_TEST_UP_SSW : BOOL ;	//FL Elevator UP PB
   HMI_ROLLER_TEST_FWD_SSW : BOOL ;	//FL Roller FWD SW
   HMI_ROLLER_TEST_REV_SSW : BOOL ;	//FL Roller REV SW
   HMI_PUSHER_1_TEST_SSW : BOOL ;	//FL Pusher 1 SW
   HMI_CONVEYOR_1_TEST_SSW : BOOL ;	//FL Conv 1 SW
   HMI_CONVEYOR_2B_TEST_SSW : BOOL ;	//FL Conv 2 Belt SW
   HMI_CONVEYOR_2L_TEST_SSW : BOOL ;	//FL Conv 2 Lift SW
   HMI_CONVEYOR_2R_TEST_SSW : BOOL ;	//FL Conv 2 Roller SW
   HMI_CONVEYOR_3_TEST_SSW : BOOL ;	//FL Conv 3 SW
   HMI_CONVEYOR_4_TEST_SSW : BOOL ;	//FL Conv 4 SW
   HMI_CONVEYOR_5_TEST_SSW : BOOL ;	//FL Conv 5 SW
   HMI_CONVEYOR_6_TEST_SSW : BOOL ;	//FL Conv 6 SW
   HMI_CONVEYOR_7_TEST_SSW : BOOL ;	//FL Flipper Conv 7 SW
   HMI_CONVEYOR_8_TEST_SSW : BOOL ;	//FL Turn Table Conv 8 SW
   HMI_TURNTABLE_CCW_SSW : BOOL ;	//FL Turn Table / Conveyor CCW PB
   HMI_TURNTABLE_CW_SSW : BOOL ;	//FL Turn Table / Conveyor CW PB
   HMI_FLIPPER_SERVICE_SSW : BOOL ;	//FL Flipper Service SW
   HMI_FLIPPER_FLIP_SSW : BOOL ;	//FL Flipper - Flip PB
   HMI_CONVEYOR_9_TEST_SSW : BOOL ;	//FL Conv 9 SW
   HMI_PUSHER_2_TEST_SSW : BOOL ;	//FL Pusher 2 SW
   HMI_PIVOT_SERVICE_SSW : BOOL ;	//FL Conv 10 - Pivot Service SW
   HMI_PIVOT_TEST_DN_SSW : BOOL ;	//FL Conv 10 - Pivot DN PB
   HMI_PIVOT_TEST_UP_SSW : BOOL ;	//FL Conv 10 - Pivot UP PB
   BIT202 : BOOL ;	//FL Spare
   BIT203 : BOOL ;	//FL Spare
   TURNTABLE_SERVICE_PBSHOW : BOOL ;	//FL TurnTable Service PB SHOW
   TURNTABLE_SERVICE_SSW : BOOL ;	//FL TurnTable Service SW
   HMI_CONVEYOR_10_TEST_SSW : BOOL ;	//FL Conv 10 - Conveyor SW
   LOADER_FING_SERVICE_SSW : BOOL ;	//FL Loader Service SW - Fingers
   LOADER_LIFT_SERVICE_SSW : BOOL ;	//FL Loader Service SW - Lift
   LOADER_LIFT_TOP_PB : BOOL ;	//FL Loader Lift - TOP PB
   LOADER_LIFT_UP_PB : BOOL ;	//FL Loader Lift - UP PB
   LOADER_LIFT_DN_PB : BOOL ;	//FL Loader Lift - DOWN PB
   FINGER_RETRACT_TEST_PB : BOOL ;	//FL Loader Fingers Retract PB
   FINGER_EXTEND_TEST_PB : BOOL ;	//FL Loader Fingers Extend PB
   FINGER_TILT_TEST_PB : BOOL ;	//FL Loader Fingers Tilt Down PB
   FINGER_BELT_TEST_SW : BOOL ;	//FL Loader Fingers Belt SW
   HMI_CONVEYOR_11_TEST_SSW : BOOL ;	//FL Conv 11 Test SW
   HMI_CONVEYOR_12_TEST_SSW : BOOL ;	//FL Conv 12 Test SW
   HMI_CONVEYOR_13_TEST_SSW : BOOL ;	//FL Conv 13 Test SW
   HMI_CONVEYOR_21_TEST_SSW : BOOL ;	//FL Conv 21 Test SW
   HMI_CONVEYOR_22_TEST_SSW : BOOL ;	//FL Conv 22 Test SW
   HMI_CONVEYOR_23_TEST_SSW : BOOL ;	//FL Conv 23 Test SW
   CONVEYOR_0_MOTOR_STATUS : BOOL ;	//FL Conveyor 0 - Motor M62.0 Status Bit
   PUSHER_0_MOTOR_STATUS : BOOL ;	//FL Pusher 0 - Motor M62.2 Status Bit
   PUSHER_0_COLOR_WORD : WORD ;	//WD Pusher 0 - 2145 - Motor Status Color
   CONV_0_COLOR_WORD : WORD ;	//WD Conveyor 0 - 2145 - Motor Status Color
   ELEVATOR_COLOR_WORD : WORD ;	//WD Elevator - Motor Status Color
   PUSHER_1_COLOR_WORD : WORD ;	//WD Pusher 1 - Motor Status Color
   CONV_1_COLOR_WORD : WORD ;	//WD Conv 1 - Motor Status Color
   CONV_2_BELT_COLOR_WORD : WORD ;	//WD Conv 2 Belt - Motor Status Color
   LIFT_ROLLER_2_COLOR_WORD : WORD ;	//WD Lift 2 Roller - Actuator Status Color
   CONV_2_ROLLER_COLOR_WORD : WORD ;	//WD Conv 2 Roller - Motor Status Color
   CONV_3_COLOR_WORD : WORD ;	//WD Conveyor 3 - Motor Status Color
   CONV_4_COLOR_WORD : WORD ;	//WD Conveyor 4 - Motor Status Color
   CONV_5_COLOR_WORD : WORD ;	//WD Conveyor 5 - Motor Status Color
   CONV_6_COLOR_WORD : WORD ;	//WD Conveyor 6 - Motor Status Color
   CONV_7_COLOR_WORD : WORD ;	//WD Conveyor 7 - Motor Status Color
   FLIPPER_COLOR_WORD : WORD ;	//WD WDipper - Motor M46.0 Status Color
   CONV_8_COLOR_WORD : WORD ;	//WD Conveyor 8 - Motor M46.4 Status Color
   TURN_TABLE_COLOR_WORD : WORD ;	//WD TurnTable - Motor M47.0 Status Color
   CONV_9_COLOR_WORD : WORD ;	//WD Conveyor 9 - Motor M47.5 Status Color
   PUSHER_2_COLOR_WORD : WORD ;	//WD Pusher 2 - Motor M47.6 Status Color
   CONV_10_COLOR_WORD : WORD ;	//WD Conveyor 10 - Motor M48.0 Status Color
   CONV_11_COLOR_WORD : WORD ;	//WD Conveyor 11 - Motor M48.3 Status Color
   CONV_12_COLOR_WORD : WORD ;	//WD Conveyor 12 - Motor M48.6 Status Color
   CONV_13_COLOR_WORD : WORD ;	//WD Conveyor 13 - Motor M49.0 Status Color
   CONV_21_COLOR_WORD : WORD ;	//WD Conveyor 21 - Motor M53.4 Status Color
   CONV_22_COLOR_WORD : WORD ;	//WD Conveyor 22 - Motor M53.6 Status Color
   CONV_23_COLOR_WORD : WORD ;	//WD Conveyor 23 - Motor M54.0 Status Color
   LOADER_LIFT_COLOR_WORD : WORD ;	//WD Loader Lift - Motor M54.6 Status Color
   LOADER_FING_COLOR_WORD : WORD ;	//WD Loader Fingers - Motor M50.5 Status Color
   FINGERS_BELT_COLOR_WORD : WORD ;	//WD Fingers Belt - Motor M54.6 Status Color
   HIGH_LEVEL_23_GRAPHIC : WORD ;	//WD High Level Conveyor 23
   LOW_LEVEL_13_GRAPHIC : WORD ;	//WD Low Level Conveyor 13
   PIVOT_GRAPHIC : WORD ;	//WD Pivot Conveyor Graphic
   CONV_3_COUNT : WORD ;	//WD Slat Conveyor 3 - Packet Count
   CONV_4_COUNT : WORD ;	//WD Collator Conveyor 4 - Packet Count
   CONV_5_COUNT : WORD ;	//WD Link Conveyor 5 - Packet Count
   CONV_6_COUNT : WORD ;	//WD Delivery Conveyor 6 - Packet Count
   CONV_10_COUNT : WORD ;	//WD Pivot Conveyor 10 - Packet Count
   CONV_11_COUNT : WORD ;	//WD Cumul Conveyor 11 - Packet Count
   CONV_12_COUNT : WORD ;	//WD Cumul Conveyor 12 - Packet Count
   CONV_13_COUNT : WORD ;	//WD Delivery Conveyor 13 - Packet Count
   CONV_21_COUNT : WORD ;	//WD Cumul Conveyor 21 - Packet Count
   CONV_22_COUNT : WORD ;	//WD Cumul Conveyor 22 - Packet Count
   CONV_23_COUNT : WORD ;	//WD Delivery Conveyor 23 - Packet Count
   FLIPPER_CCW : WORD ;	//WD Flipper Graphic CCW
   FLIPPER_CW : WORD ;	//WD Flipper Graphic CW
   FLIPPER_POSITION : WORD ;	//WD Flipper Positioning mS
   TURN_COLOR : WORD ;	//WD Turn Table - Turn Color
   FLIPPER_COLOR : WORD ;	//WD Flipper Color
   FLIPPER_PACK_PRESENCE : WORD ;	//WD Flipper - Packet Presence
   TURNTABLE_PACK_PRESENCE : WORD ;	//WD TurnTable - Packet Presence
   ROLLER_PACK_PRESENCE : WORD ;	//WD Pusher Roller - Packet Presence
   PUSHER_PACK_PRESENCE : WORD ;	//WD Pusher - Packet Presence
   CONV_0_STATUS : BOOL ;	//FL Conveyor 0 - Motor Status Bit
   PUSHER_0_STATUS : BOOL ;	//FL Pusher 0 - Motor Status
   ELEVATOR_STATUS : BOOL ;	//FL Elevator - Motor Status
   PUSHER_1_STATUS : BOOL ;	//FL Pusher 1 - Motor Status
   CONV_1_STATUS : BOOL ;	//FL Conveyor 1 - Motor Status
   TURNTABLE_RNDTRIP : BOOL ;	//FL TurnTable Round Trip CMD
   RNDTRIP_PB_VISIBLE : BOOL ;	//FL TurnTable Round Trip PB Visible
   BOOL_SPARE227 : BOOL ;	//FL
   SCREEN_CALL_0 : BOOL ;	//FL  HMI Call Screen 0
   SCREEN_CALL_1 : BOOL ;	//FL  HMI Call Screen 1
   SCREEN_CALL_2 : BOOL ;	//FL  HMI Call Screen 2
   SCREEN_CALL_3 : BOOL ;	//FL  HMI Call Screen 3
   SCREEN_CALL_4 : BOOL ;	//FL  HMI Call Screen 4
   BOOL_SPARE2276 : BOOL ;	//FL
   BOOL_SPARE2277 : BOOL ;	//FL
   BOOL_SPARE2278 : BOOL ;	//FL
   BOOL_SPARE2279 : BOOL ;	//FL
   BOOL_SPARE22710 : BOOL ;	//FL
   BOOL_SPARE22711 : BOOL ;	//FL
   BOOL_SPARE22712 : BOOL ;	//FL
   BOOL_SPARE22713 : BOOL ;	//FL
   BOOL_SPARE22714 : BOOL ;	//FL
   BOOL_SPARE22715 : BOOL ;	//FL
   BOOL_SPARE22716 : BOOL ;	//FL
   BOOL_SPARE22717 : BOOL ;	//FL
   BOOL_SPARE22718 : BOOL ;	//FL
   BOOL_SPARE22719 : BOOL ;	//FL
   BOOL_SPARE22720 : BOOL ;	//FL
   BOOL_SPARE22721 : BOOL ;	//FL
   BOOL_SPARE22722 : BOOL ;	//FL
   BOOL_SPARE22723 : BOOL ;	//FL
   BOOL_SPARE22724 : BOOL ;	//FL
   WORD_SPARE23 : WORD ;	//WD
   FLIPPER_TURN_COLOR : WORD ;	//WD Flipper Turn Color
   NEW_ORDER_COLOR : WORD ;	//WD Conveyor 10 - New Order Color
   SERVICE_FLIPPER : BOOL ;	//FLS Flipper Service - Switch
   FLIP_TEST : BOOL ;	//FLS Flipper Flip - Test Switch
   SERVICE_TURNTABLE : BOOL ;	//FLS TurnTable Service - Switch
   TURN_TEST_CW : BOOL ;	//FLS TurnTable - Turn CW - Status Bit
   TURN_TEST_CCW : BOOL ;	//FLS TurnTable - Turn CCW - Status Bit
   PUSHER_2_TEST : BOOL ;	//FLS Pusher 2 - Test Switch
   CONVEYOR_10_TEST_SW : BOOL ;	//FLS Collator Conveyor 10 - Test Switch
   PIVOT_SERVICE_SW : BOOL ;	//FL Pivot Service - Status
   PIVOT_UP_TEST_PB : BOOL ;	//FLS Pivot Conveyor UP - Test Switch
   PIVOT_DN_TEST_PB : BOOL ;	//FLS Pivot Conveyor DN - Test Switch
   PIVOT_STATUS : BOOL ;	//FL Pivot ON - Status
   CONV_8_INVERT_SELECT : BOOL ;	//FL TurnTable Conveyor 8 - Positioning Time - Display Selector Bit - INVERT
   CONVEYOR_11_TEST_SW : BOOL ;	//FLS Cumul Conveyor 11 - Test Switch
   CONVEYOR_12_TEST_SW : BOOL ;	//FLS Cumul Conveyor 12 - Test Switch
   CONVEYOR_13_TEST_SW : BOOL ;	//FLS Delivery Conveyor 13 - Test Switch
   CONVEYOR_21_TEST_SW : BOOL ;	//FLS Cumul Conveyor 21 - Test Switch
   CONVEYOR_22_TEST_SW : BOOL ;	//FLS Cumul Conveyor 22 - Test Switch
   CONVEYOR_23_TEST_SW : BOOL ;	//FLS Delivery Conveyor 23 - Test Switch
   LOADER_SERVICE_SW : BOOL ;	//FLS Loader Service - Switch
   LOADER_UP_TEST_PB : BOOL ;	//FLS Loader Lift Up - Test Switch
   LOADER_DN_TEST_PB : BOOL ;	//FLS Loader Lift Dn - Test Switch
   FINGERS_EXTEND_TEST_PB : BOOL ;	//FLS Loader Finger Extend - Test Switch
   FINGERS_RETRACT_TEST_PB : BOOL ;	//FLS Loader Finger Retract - Test Switch
   FP_ONESHOT_0 : BOOL ;	//FP One Shot
   CONVEYOR_0_SERVICE_SW : BOOL ;	//FL Conveyor 0 / Pusher 0 - Service Enable
   ELEVATOR_SERVICE_SW : BOOL ;	//FL Elevator / Pusher 1 - Service Enable
   CONVEYOR_1_SERVICE_SW : BOOL ;	//FL Conveyor 1 - Service Enable Select - Screen 4
   CONVEYOR_2_SERVICE_SW : BOOL ;	//FL Conveyor 2 - Service Enable Select - Screen 4
   CONVEYOR_3_SERVICE_SW : BOOL ;	//FL Conveyor 3 - Service Enable Select - Screen 4
   CONVEYOR_4_SERVICE_SW : BOOL ;	//FL Conveyor 4 - Service Enable Select - Screen 4
   CONVEYOR_5_SERVICE_SW : BOOL ;	//FL Conveyor 5 - Service Enable Select - Screen 4
   CONVEYOR_6_SERVICE_SW : BOOL ;	//FL Conveyor 6 - Service Enable Select - Screen 4
   CONVEYOR_7_SERVICE_SW : BOOL ;	//FL Conveyor 7 / Flipper - Service Enable Select - Screen 4
   CONVEYOR_8_SERVICE_SW : BOOL ;	//FL Conveyor 8 / TurnTable - Service Enable Select - Screen 4
   CONVEYOR_9_SERVICE_SW : BOOL ;	//FL Conveyor 9 / Pusher 2 - Service Enable Select - Screen 4
   CONVEYOR_10_SERVICE_SW : BOOL ;	//FL Conveyor 10 - Service Enable Select - Screen 4
   CONVEYOR_11_SERVICE_SW : BOOL ;	//FL Conveyors 11, 12, 13 - Service Enable Select - Screen 4
   CONVEYOR_21_SERVICE_SW : BOOL ;	//FL Conveyors 21, 22, 23 - Service Enable Select - Screen 4
   LOADER_SERVICE_ENABLE_SW : BOOL ;	//FL Loader - Service Enable
   CTRL48 : BOOL ;	//FL Spare - Service Enable
   CTRL49 : BOOL ;	//FL Spare -
   CTRL50 : BOOL ;	//FL Spare -
   CTRL51 : BOOL ;	//FL Spare -
   CTRL52 : BOOL ;	//FL Spare -
   CTRL53 : BOOL ;	//FL Spare -
   CTRL54 : BOOL ;	//FL Spare -
   CTRL55 : BOOL ;	//FL Spare -
   CTRL56 : BOOL ;	//FL Spare -
   CLEARING_FUNCTION : WORD ;	//WD Clearing Function - Underneat Rectangle
   WORD57 : WORD ;	//WD
   WORD58 : WORD ;	//WD
   ACTUAL_HMI_SCREEN_NO : WORD ;	//WD HMI Actual Display Screen
   CONVEYOR_MAXCOUNT_L : WORD  := W#16#6;	//WD All Conveyors Max Count Lenght (6)
   CONVEYOR_MAXCOUNT_W : WORD  := W#16#7;	//WD All Conveyors Max Count Widtht (7)
   WORD62 : WORD ;	//WD
   CONV_7_POS_mS : WORD ;	//WD Flipper Conveyor 7 - Positioning Time x10 [mS]
   CONV_8_POS_FWD_mS : WORD ;	//WD TurnTable Conveyor 8 - FWD Positioning Time x10 [mS]
   CONV_8_POS_REV_mS : WORD ;	//WD TurnTable Conveyor 8 - REV Positioning Time x10 [mS]
   CONV_9_POS_mS : WORD ;	//WD Pusher 2 Conveyor 9 - Positioning Time x10 [mS]
   WORD_PACKET_LENGTH : WORD ;	//WD Actual Packet Length mm
   DELAY_DISPLAY_7 : WORD ;	//WD HMI Flipper 7 Delay Display
   DELAY_DISPLAY_9 : WORD ;	//WD HMI Conveyor 9 Delay Display
   WORD_SPARE2 : WORD ;
   WORD_SPARE3 : WORD ;
   WORD_SPARE4 : WORD ;
  END_STRUCT ;
BEGIN
   GRAPHIC_INIT := FALSE;
   EMERGENCY_BLINK := FALSE;
   TRANS_SYSTEM_ON_SW := FALSE;
   COMPRESSED_AIR := FALSE;
   TRANS_SYSTEM_RUN_STATUS := FALSE;
   PACKET_in_FLIPPER_SW := FALSE;
   SERVICE_INIT_PB := FALSE;
   ALL_SERVICE_ENABLE_SW := FALSE;
   SERVICE_SW_1_STATUS := FALSE;
   SERVICE_SW_2_STATUS := FALSE;
   SERVICE_SW_3_STATUS := FALSE;
   SERVICE_SW_1_2_STATUS := FALSE;
   BIT12 := FALSE;
   BIT13 := FALSE;
   SERVICE_SW_2_TIME_ADJ := FALSE;
   PACKETIZER_GATE_STATUS := FALSE;
   E_STOP_CONSOLE_STATUS := FALSE;
   E_STOP_ELEVATOR_STATUS := FALSE;
   E_STOP_FLIPPER_STATUS := FALSE;
   E_STOP_LOADER_STATUS := FALSE;
   HAND_FEED_ARROW_STATUS := FALSE;
   ELEVATOR_DOOR_STATUS := FALSE;
   FLIPPER_DOOR_STATUS := FALSE;
   LOADER_DOOR_STATUS := FALSE;
   LIGHT_BARRIER_1_STATUS := FALSE;
   LIGHT_BARRIER_2_STATUS := FALSE;
   LIGHT_BARRIER_3_STATUS := FALSE;
   LIGHT_BARRIER_4_STATUS := FALSE;
   LIGHT_BARRIER_5_STATUS := FALSE;
   LIGHT_BARRIER_6_STATUS := FALSE;
   LIGHT_BARRIER_B_STATUS := FALSE;
   LIGHT_BARRIER_A_STATUS := FALSE;
   BIT32 := FALSE;
   BIT33 := FALSE;
   BIT34 := FALSE;
   BIT35 := FALSE;
   BIT36 := FALSE;
   BIT37 := FALSE;
   BIT38 := FALSE;
   BIT39 := FALSE;
   BIT40 := FALSE;
   BIT41 := FALSE;
   BIT42 := FALSE;
   BIT43 := FALSE;
   BIT44 := FALSE;
   BIT45 := FALSE;
   BIT46 := FALSE;
   BIT47 := FALSE;
   BIT48 := FALSE;
   BIT49 := FALSE;
   BIT50 := FALSE;
   BIT51 := FALSE;
   BIT52 := FALSE;
   BIT53 := FALSE;
   BIT54 := FALSE;
   BIT55 := FALSE;
   BIT56 := FALSE;
   BIT57 := FALSE;
   BIT58 := FALSE;
   BIT59 := FALSE;
   BIT60 := FALSE;
   BIT61 := FALSE;
   BIT62 := FALSE;
   CONVEYORS_CLEARING := FALSE;
   ELEVATOR_MOTOR_STATUS := FALSE;
   PUSHER_1_MOTOR_STATUS := FALSE;
   CONVEYOR_1_MOTOR_STATUS := FALSE;
   CONVEYOR_2B_MOTOR_STATUS := FALSE;
   CONVEYOR_2R_MOTOR_STATUS := FALSE;
   CONVEYOR_3_MOTOR_STATUS := FALSE;
   CONVEYOR_4_MOTOR_STATUS := FALSE;
   CONVEYOR_5_MOTOR_STATUS := FALSE;
   CONVEYOR_6_MOTOR_STATUS := FALSE;
   CONVEYOR_7_MOTOR_STATUS := FALSE;
   FLIPPER_MOTOR_STATUS := FALSE;
   CONVEYOR_8_MOTOR_STATUS := FALSE;
   TURNTABLE_MOTOR_STATUS := FALSE;
   CONVEYOR_9_MOTOR_STATUS := FALSE;
   PUSHER_2_MOTOR_STATUS := FALSE;
   CONVEYOR_10_MOTOR_STATUS := FALSE;
   CONVEYOR_11_MOTOR_STATUS := FALSE;
   CONVEYOR_12_MOTOR_STATUS := FALSE;
   CONVEYOR_13_MOTOR_STATUS := FALSE;
   CONVEYOR_21_MOTOR_STATUS := FALSE;
   CONVEYOR_22_MOTOR_STATUS := FALSE;
   CONVEYOR_23_MOTOR_STATUS := FALSE;
   LOADER_LIFT_MOTOR_STATUS := FALSE;
   LOADER_FING_MOTOR_STATUS := FALSE;
   LOADER_BELT_MOTOR_STATUS := FALSE;
   LIGHT_BARRIER_7_STATUS := FALSE;
   LIGHT_BARRIER_8_STATUS := FALSE;
   LIGHT_BARRIER_9_STATUS := FALSE;
   LIGHT_BARRIER_10_STATUS := FALSE;
   LIGHT_BARRIER_11_STATUS := FALSE;
   LIGHT_BARRIER_12_STATUS := FALSE;
   LIGHT_BARRIER_13_STATUS := FALSE;
   LIGHT_BARRIER_14_STATUS := FALSE;
   LIGHT_BARRIER_15_STATUS := FALSE;
   LIGHT_BARRIER_16_STATUS := FALSE;
   LIGHT_BARRIER_17_STATUS := FALSE;
   LIGHT_BARRIER_18_STATUS := FALSE;
   LIGHT_BARRIER_19_STATUS := FALSE;
   LIGHT_BARRIER_20_STATUS := FALSE;
   LIGHT_BARRIER_21_STATUS := FALSE;
   LIGHT_BARRIER_22_STATUS := FALSE;
   LIGHT_BARRIER_23_STATUS := FALSE;
   LIGHT_BARRIER_24_STATUS := FALSE;
   LIGHT_BARRIER_25_STATUS := FALSE;
   LIGHT_BARRIER_26_STATUS := FALSE;
   LIGHT_BARRIER_27_STATUS := FALSE;
   LIGHT_BARRIER_28_STATUS := FALSE;
   LIGHT_BARRIER_29_STATUS := FALSE;
   LIGHT_BARRIER_30_STATUS := FALSE;
   LIGHT_BARRIER_31_STATUS := FALSE;
   LIGHT_BARRIER_32_STATUS := FALSE;
   PROX_9_STATUS := FALSE;
   PROX_10_STATUS := FALSE;
   PROX_11_STATUS := FALSE;
   PROX_12_STATUS := FALSE;
   PROX_13_STATUS := FALSE;
   PROX_14_STATUS := FALSE;
   PROX_15_STATUS := FALSE;
   PROX_16_STATUS := FALSE;
   PROX_17_STATUS := FALSE;
   PROX_18_STATUS := FALSE;
   PROX_19_STATUS := FALSE;
   PROX_20_STATUS := FALSE;
   PROX_21_STATUS := FALSE;
   PROX_22_STATUS := FALSE;
   PROX_23_STATUS := FALSE;
   PROX_24_STATUS := FALSE;
   FP131 := FALSE;
   FP132 := FALSE;
   FP133 := FALSE;
   FP134 := FALSE;
   FP135 := FALSE;
   TURNTABLE_DELIV_POSITION := FALSE;
   TURNTABLE_REVERSE_ARROW := FALSE;
   TURNTABLE_DIR_SELECT_SW := FALSE;
   TURNTABLE_FLICK_MOTION := FALSE;
   FP140 := FALSE;
   FP141 := FALSE;
   FP142 := FALSE;
   FP143 := FALSE;
   PROX_1_STATUS := FALSE;
   PROX_2_STATUS := FALSE;
   PROX_3_STATUS := FALSE;
   PROX_4_STATUS := FALSE;
   PROX_5_STATUS := FALSE;
   PROX_6_STATUS := FALSE;
   PROX_7_STATUS := FALSE;
   PROX_8_STATUS := FALSE;
   BIT152 := FALSE;
   BIT153 := FALSE;
   BIT154 := FALSE;
   BIT155 := FALSE;
   BIT156 := FALSE;
   BIT157 := FALSE;
   BIT158 := FALSE;
   BIT159 := FALSE;
   SERVICE_SSW_MAIN := FALSE;
   SERVICE_SSW_STATUS := FALSE;
   CLEARING_SSW_MAIN := FALSE;
   CLEARING_SSW_STATUS := FALSE;
   MAN_FEED_SSW_MAIN := FALSE;
   MAN_FEED_SSW_STATUS := FALSE;
   TURNTABLE_SSW_MAIN := FALSE;
   TURNTABLE_SSW_STATUS := FALSE;
   FLIPPER_SSW_MAIN := FALSE;
   FLIPPER_SSW_STATUS := FALSE;
   ROLLER_SSW_MAIN := FALSE;
   ROLLER_SSW_STATUS := FALSE;
   ELEVATOR_ROUND_TRIP_SSW := FALSE;
   BIT173 := FALSE;
   BIT174 := FALSE;
   BIT175 := FALSE;
   HMI_PUSHER_0_TEST_SSW := FALSE;
   HMI_ELEVATOR_SERVICE_SSW := FALSE;
   HMI_ELEVATOR_TEST_DN_SSW := FALSE;
   HMI_ELEVATOR_TEST_UP_SSW := FALSE;
   HMI_ROLLER_TEST_FWD_SSW := FALSE;
   HMI_ROLLER_TEST_REV_SSW := FALSE;
   HMI_PUSHER_1_TEST_SSW := FALSE;
   HMI_CONVEYOR_1_TEST_SSW := FALSE;
   HMI_CONVEYOR_2B_TEST_SSW := FALSE;
   HMI_CONVEYOR_2L_TEST_SSW := FALSE;
   HMI_CONVEYOR_2R_TEST_SSW := FALSE;
   HMI_CONVEYOR_3_TEST_SSW := FALSE;
   HMI_CONVEYOR_4_TEST_SSW := FALSE;
   HMI_CONVEYOR_5_TEST_SSW := FALSE;
   HMI_CONVEYOR_6_TEST_SSW := FALSE;
   HMI_CONVEYOR_7_TEST_SSW := FALSE;
   HMI_CONVEYOR_8_TEST_SSW := FALSE;
   HMI_TURNTABLE_CCW_SSW := FALSE;
   HMI_TURNTABLE_CW_SSW := FALSE;
   HMI_FLIPPER_SERVICE_SSW := FALSE;
   HMI_FLIPPER_FLIP_SSW := FALSE;
   HMI_CONVEYOR_9_TEST_SSW := FALSE;
   HMI_PUSHER_2_TEST_SSW := FALSE;
   HMI_PIVOT_SERVICE_SSW := FALSE;
   HMI_PIVOT_TEST_DN_SSW := FALSE;
   HMI_PIVOT_TEST_UP_SSW := FALSE;
   BIT202 := FALSE;
   BIT203 := FALSE;
   TURNTABLE_SERVICE_PBSHOW := FALSE;
   TURNTABLE_SERVICE_SSW := FALSE;
   HMI_CONVEYOR_10_TEST_SSW := FALSE;
   LOADER_FING_SERVICE_SSW := FALSE;
   LOADER_LIFT_SERVICE_SSW := FALSE;
   LOADER_LIFT_TOP_PB := FALSE;
   LOADER_LIFT_UP_PB := FALSE;
   LOADER_LIFT_DN_PB := FALSE;
   FINGER_RETRACT_TEST_PB := FALSE;
   FINGER_EXTEND_TEST_PB := FALSE;
   FINGER_TILT_TEST_PB := FALSE;
   FINGER_BELT_TEST_SW := FALSE;
   HMI_CONVEYOR_11_TEST_SSW := FALSE;
   HMI_CONVEYOR_12_TEST_SSW := FALSE;
   HMI_CONVEYOR_13_TEST_SSW := FALSE;
   HMI_CONVEYOR_21_TEST_SSW := FALSE;
   HMI_CONVEYOR_22_TEST_SSW := FALSE;
   HMI_CONVEYOR_23_TEST_SSW := FALSE;
   CONVEYOR_0_MOTOR_STATUS := FALSE;
   PUSHER_0_MOTOR_STATUS := FALSE;
   PUSHER_0_COLOR_WORD := W#16#0;
   CONV_0_COLOR_WORD := W#16#0;
   ELEVATOR_COLOR_WORD := W#16#3226;
   PUSHER_1_COLOR_WORD := W#16#0;
   CONV_1_COLOR_WORD := W#16#0;
   CONV_2_BELT_COLOR_WORD := W#16#0;
   LIFT_ROLLER_2_COLOR_WORD := W#16#0;
   CONV_2_ROLLER_COLOR_WORD := W#16#0;
   CONV_3_COLOR_WORD := W#16#0;
   CONV_4_COLOR_WORD := W#16#0;
   CONV_5_COLOR_WORD := W#16#0;
   CONV_6_COLOR_WORD := W#16#0;
   CONV_7_COLOR_WORD := W#16#0;
   FLIPPER_COLOR_WORD := W#16#0;
   CONV_8_COLOR_WORD := W#16#0;
   TURN_TABLE_COLOR_WORD := W#16#0;
   CONV_9_COLOR_WORD := W#16#0;
   PUSHER_2_COLOR_WORD := W#16#0;
   CONV_10_COLOR_WORD := W#16#0;
   CONV_11_COLOR_WORD := W#16#0;
   CONV_12_COLOR_WORD := W#16#0;
   CONV_13_COLOR_WORD := W#16#0;
   CONV_21_COLOR_WORD := W#16#0;
   CONV_22_COLOR_WORD := W#16#0;
   CONV_23_COLOR_WORD := W#16#0;
   LOADER_LIFT_COLOR_WORD := W#16#0;
   LOADER_FING_COLOR_WORD := W#16#0;
   FINGERS_BELT_COLOR_WORD := W#16#0;
   HIGH_LEVEL_23_GRAPHIC := W#16#0;
   LOW_LEVEL_13_GRAPHIC := W#16#0;
   PIVOT_GRAPHIC := W#16#0;
   CONV_3_COUNT := W#16#0;
   CONV_4_COUNT := W#16#0;
   CONV_5_COUNT := W#16#0;
   CONV_6_COUNT := W#16#0;
   CONV_10_COUNT := W#16#0;
   CONV_11_COUNT := W#16#0;
   CONV_12_COUNT := W#16#0;
   CONV_13_COUNT := W#16#4;
   CONV_21_COUNT := W#16#0;
   CONV_22_COUNT := W#16#0;
   CONV_23_COUNT := W#16#0;
   FLIPPER_CCW := W#16#0;
   FLIPPER_CW := W#16#0;
   FLIPPER_POSITION := W#16#0;
   TURN_COLOR := W#16#0;
   FLIPPER_COLOR := W#16#0;
   FLIPPER_PACK_PRESENCE := W#16#0;
   TURNTABLE_PACK_PRESENCE := W#16#0;
   ROLLER_PACK_PRESENCE := W#16#0;
   PUSHER_PACK_PRESENCE := W#16#0;
   CONV_0_STATUS := FALSE;
   PUSHER_0_STATUS := FALSE;
   ELEVATOR_STATUS := FALSE;
   PUSHER_1_STATUS := FALSE;
   CONV_1_STATUS := FALSE;
   TURNTABLE_RNDTRIP := FALSE;
   RNDTRIP_PB_VISIBLE := FALSE;
   BOOL_SPARE227 := FALSE;
   SCREEN_CALL_0 := FALSE;
   SCREEN_CALL_1 := FALSE;
   SCREEN_CALL_2 := FALSE;
   SCREEN_CALL_3 := FALSE;
   SCREEN_CALL_4 := FALSE;
   BOOL_SPARE2276 := FALSE;
   BOOL_SPARE2277 := FALSE;
   BOOL_SPARE2278 := FALSE;
   BOOL_SPARE2279 := FALSE;
   BOOL_SPARE22710 := FALSE;
   BOOL_SPARE22711 := FALSE;
   BOOL_SPARE22712 := FALSE;
   BOOL_SPARE22713 := FALSE;
   BOOL_SPARE22714 := FALSE;
   BOOL_SPARE22715 := FALSE;
   BOOL_SPARE22716 := FALSE;
   BOOL_SPARE22717 := FALSE;
   BOOL_SPARE22718 := FALSE;
   BOOL_SPARE22719 := FALSE;
   BOOL_SPARE22720 := FALSE;
   BOOL_SPARE22721 := FALSE;
   BOOL_SPARE22722 := FALSE;
   BOOL_SPARE22723 := FALSE;
   BOOL_SPARE22724 := FALSE;
   WORD_SPARE23 := W#16#0;
   FLIPPER_TURN_COLOR := W#16#0;
   NEW_ORDER_COLOR := W#16#0;
   SERVICE_FLIPPER := FALSE;
   FLIP_TEST := FALSE;
   SERVICE_TURNTABLE := FALSE;
   TURN_TEST_CW := FALSE;
   TURN_TEST_CCW := FALSE;
   PUSHER_2_TEST := FALSE;
   CONVEYOR_10_TEST_SW := FALSE;
   PIVOT_SERVICE_SW := FALSE;
   PIVOT_UP_TEST_PB := FALSE;
   PIVOT_DN_TEST_PB := FALSE;
   PIVOT_STATUS := FALSE;
   CONV_8_INVERT_SELECT := FALSE;
   CONVEYOR_11_TEST_SW := FALSE;
   CONVEYOR_12_TEST_SW := FALSE;
   CONVEYOR_13_TEST_SW := FALSE;
   CONVEYOR_21_TEST_SW := FALSE;
   CONVEYOR_22_TEST_SW := FALSE;
   CONVEYOR_23_TEST_SW := FALSE;
   LOADER_SERVICE_SW := FALSE;
   LOADER_UP_TEST_PB := FALSE;
   LOADER_DN_TEST_PB := FALSE;
   FINGERS_EXTEND_TEST_PB := FALSE;
   FINGERS_RETRACT_TEST_PB := FALSE;
   FP_ONESHOT_0 := FALSE;
   CONVEYOR_0_SERVICE_SW := FALSE;
   ELEVATOR_SERVICE_SW := FALSE;
   CONVEYOR_1_SERVICE_SW := FALSE;
   CONVEYOR_2_SERVICE_SW := FALSE;
   CONVEYOR_3_SERVICE_SW := FALSE;
   CONVEYOR_4_SERVICE_SW := FALSE;
   CONVEYOR_5_SERVICE_SW := FALSE;
   CONVEYOR_6_SERVICE_SW := FALSE;
   CONVEYOR_7_SERVICE_SW := FALSE;
   CONVEYOR_8_SERVICE_SW := FALSE;
   CONVEYOR_9_SERVICE_SW := FALSE;
   CONVEYOR_10_SERVICE_SW := FALSE;
   CONVEYOR_11_SERVICE_SW := FALSE;
   CONVEYOR_21_SERVICE_SW := FALSE;
   LOADER_SERVICE_ENABLE_SW := FALSE;
   CTRL48 := FALSE;
   CTRL49 := FALSE;
   CTRL50 := FALSE;
   CTRL51 := FALSE;
   CTRL52 := FALSE;
   CTRL53 := FALSE;
   CTRL54 := FALSE;
   CTRL55 := FALSE;
   CTRL56 := FALSE;
   CLEARING_FUNCTION := W#16#0;
   WORD57 := W#16#0;
   WORD58 := W#16#0;
   ACTUAL_HMI_SCREEN_NO := W#16#0;
   CONVEYOR_MAXCOUNT_L := W#16#6;
   CONVEYOR_MAXCOUNT_W := W#16#7;
   WORD62 := W#16#0;
   CONV_7_POS_mS := W#16#96;
   CONV_8_POS_FWD_mS := W#16#0;
   CONV_8_POS_REV_mS := W#16#0;
   CONV_9_POS_mS := W#16#0;
   WORD_PACKET_LENGTH := W#16#0;
   DELAY_DISPLAY_7 := W#16#0;
   DELAY_DISPLAY_9 := W#16#0;
   WORD_SPARE2 := W#16#0;
   WORD_SPARE3 := W#16#0;
   WORD_SPARE4 := W#16#0;
END_DATA_BLOCK

DATA_BLOCK "HMI ALARMS"
TITLE =HMI Alarms - NS12
//One BOOL per alarm, written by FC1220 every scan (no latching here: the
//fault bits keep their own latch / reset). NS12 address: SERIALA:DB0013_DBXbbbbb.ii
//v1.1 2026-11-24: DBX9.6 Any_Fault (bytes 0...8) and DBX9.7 Any_Alarm (+ status
//9.0...9.3) for the NS12 alarm bar Control Flag (bar shown only when needed).
VERSION : 1.1


  STRUCT
   Fuse_Fault : BOOL ;	//DBX0.0 Fuse fault
   Motor_Protect : BOOL ;	//DBX0.1 Motor protection tripped
   Motor_Temp : BOOL ;	//DBX0.2 Motor temperature fault
   Air_Low : BOOL ;	//DBX0.3 Compressed air below 5 bar
   EStop_Desk_X120 : BOOL ;	//DBX0.4 E-STOP desk X120 (HMI box)
   EStop_Desk_X121 : BOOL ;	//DBX0.5 E-STOP desk X121 (feeder box)
   EStop_Elevator : BOOL ;	//DBX0.6 E-STOP elevator station
   EStop_Flipper : BOOL ;	//DBX0.7 E-STOP flipper station
   Door_Feeder : BOOL ;	//DBX1.0 Door open - feeder
   Door_Elevator : BOOL ;	//DBX1.1 Door open - elevator
   Door_Flipper : BOOL ;	//DBX1.2 Door open - flipper
   Spare_1_3 : BOOL ;	//DBX1.3 Spare
   Spare_1_4 : BOOL ;	//DBX1.4 Spare
   Spare_1_5 : BOOL ;	//DBX1.5 Spare
   Spare_1_6 : BOOL ;	//DBX1.6 Spare
   Spare_1_7 : BOOL ;	//DBX1.7 Spare
   C2_Angle_Fault : BOOL ;	//DBX2.0 C2 angle conveyor fault
   Elev_Rollers_Fault : BOOL ;	//DBX2.1 Elevator rollers (C0) fault
   Elev_Pusher_Fault : BOOL ;	//DBX2.2 Elevator pusher fault
   Elev_Not_Centered : BOOL ;	//DBX2.3 Elevator - packet not centered
   C4_Fault : BOOL ;	//DBX2.4 C4 collator fault
   C4_Timeout : BOOL ;	//DBX2.5 C4 collator timeout stop
   C4_Infeed_Obstruct : BOOL ;	//DBX2.6 C4 infeed obstruction
   C6_Fault : BOOL ;	//DBX2.7 C6 flipper delivery fault
   Flipper_Obstruct : BOOL ;	//DBX3.0 Flipper flip obstructed
   C10_Fault : BOOL ;	//DBX3.1 C10 pivot conveyor fault
   Pivot_Timeout : BOOL ;	//DBX3.2 Pivot timeout
   Pivot_Conflict : BOOL ;	//DBX3.3 Pivot / conveyor conflict
   C13_Delivery_Fault : BOOL ;	//DBX3.4 C13 delivery fault (low)
   C23_Delivery_Fault : BOOL ;	//DBX3.5 C23 delivery fault (high)
   Spare_3_6 : BOOL ;	//DBX3.6 Spare
   Spare_3_7 : BOOL ;	//DBX3.7 Spare
   VFD_U44_3 : BOOL ;	//DBX4.0 Drive U44.3 fault - C4
   VFD_U45_0 : BOOL ;	//DBX4.1 Drive U45.0 fault - C5
   VFD_U45_3 : BOOL ;	//DBX4.2 Drive U45.3 fault - C6
   VFD_U45_6 : BOOL ;	//DBX4.3 Drive U45.6 fault - C7 flipper conveyor
   VFD_U46_0 : BOOL ;	//DBX4.4 Drive U46.0 fault - Flipper
   VFD_U46_4 : BOOL ;	//DBX4.5 Drive U46.4 fault - C8 turntable conveyor
   VFD_U47_0 : BOOL ;	//DBX4.6 Drive U47.0 fault - Turntable
   VFD_U47_5 : BOOL ;	//DBX4.7 Drive U47.5 fault - C9 pusher 2 conveyor
   VFD_U47_6 : BOOL ;	//DBX5.0 Drive U47.6 fault - Pusher 2
   VFD_U48_0 : BOOL ;	//DBX5.1 Drive U48.0 fault - C10
   VFD_U48_3 : BOOL ;	//DBX5.2 Drive U48.3 fault - C11
   VFD_U48_6 : BOOL ;	//DBX5.3 Drive U48.6 fault - C12
   VFD_U49_0 : BOOL ;	//DBX5.4 Drive U49.0 fault - C13
   VFD_U53_2 : BOOL ;	//DBX5.5 Drive U53.2 fault - C21
   VFD_U53_4 : BOOL ;	//DBX5.6 Drive U53.4 fault - C22
   VFD_U54_0 : BOOL ;	//DBX5.7 Drive U54.0 fault - C23
   Sens_B5_1_On : BOOL ;	//DBX6.0 Sensor Elevator platform infeed B5.1 ON - line empty (packet left or dir
   Sens_B5_2_On : BOOL ;	//DBX6.1 Sensor Elevator platform limit B5.2 ON - line empty (packet left or dirt
   Sens_B5_4_On : BOOL ;	//DBX6.2 Sensor C1 exit B5.4 ON - line empty (packet left or dirty sensor)
   Sens_B5_5_On : BOOL ;	//DBX6.3 Sensor C2 infeed B5.5 ON - line empty (packet left or dirty sensor)
   Sens_B6_0_On : BOOL ;	//DBX6.4 Sensor C2 roller center B6.0 ON - line empty (packet left or dirty senso
   Sens_B6_7_On : BOOL ;	//DBX6.5 Sensor C4 infeed B6.7 ON - line empty (packet left or dirty sensor)
   Sens_B7_0_On : BOOL ;	//DBX6.6 Sensor C4 exit B7.0 ON - line empty (packet left or dirty sensor)
   Sens_B7_1_On : BOOL ;	//DBX6.7 Sensor C5 exit B7.1 ON - line empty (packet left or dirty sensor)
   Sens_B7_2_On : BOOL ;	//DBX7.0 Sensor C6 reaching B7.2 ON - line empty (packet left or dirty sensor)
   Sens_B7_3_On : BOOL ;	//DBX7.1 Sensor C6 exit B7.3 ON - line empty (packet left or dirty sensor)
   Sens_B7_4_On : BOOL ;	//DBX7.2 Sensor Flipper infeed B7.4 ON - line empty (packet left or dirty sensor)
   Sens_B8_2_On : BOOL ;	//DBX7.3 Sensor Flipper exit B8.2 ON - line empty (packet left or dirty sensor)
   Sens_B9_6_On : BOOL ;	//DBX7.4 Sensor C9 infeed B9.6 ON - line empty (packet left or dirty sensor)
   Sens_B9_7_On : BOOL ;	//DBX7.5 Sensor C9 packet edge B9.7 ON - line empty (packet left or dirty sensor)
   Sens_B10_4_On : BOOL ;	//DBX7.6 Sensor C10 infeed B10.4 ON - line empty (packet left or dirty sensor)
   Sens_B10_5_On : BOOL ;	//DBX7.7 Sensor C10 full B10.5 ON - line empty (packet left or dirty sensor)
   Sens_B10_7_On : BOOL ;	//DBX8.0 Sensor C11 exit B10.7 ON - line empty (packet left or dirty sensor)
   Sens_B11_0_On : BOOL ;	//DBX8.1 Sensor C12 exit B11.0 ON - line empty (packet left or dirty sensor)
   Sens_B11_1_On : BOOL ;	//DBX8.2 Sensor C13 slow B11.1 ON - line empty (packet left or dirty sensor)
   Sens_B5_4_Off : BOOL ;	//DBX8.3 Sensor C1 exit B5.4 OFF - line empty (check sensor / reflector)
   Sens_B9_7_Off : BOOL ;	//DBX8.4 Sensor C9 packet edge B9.7 OFF - line empty (check sensor / reflector)
   Spare_8_5 : BOOL ;	//DBX8.5 Spare
   Spare_8_6 : BOOL ;	//DBX8.6 Spare
   Spare_8_7 : BOOL ;	//DBX8.7 Spare
   Clearing_Active : BOOL ;	//DBX9.0 Clearing (F4) active
   Packets_Present : BOOL ;	//DBX9.1 Packets present on C1-C2 / C7-C9
   Control_Off : BOOL ;	//DBX9.2 Control voltage OFF - press START
   Start_Ready : BOOL ;	//DBX9.3 Start ready (10 s)
   Spare_9_4 : BOOL ;	//DBX9.4 Spare
   Spare_9_5 : BOOL ;	//DBX9.5 Spare
   Any_Fault : BOOL ;	//DBX9.6 At Least One Fault (DBX0.0...8.7) - NS12 Alarm Bar Display
   Any_Alarm : BOOL ;	//DBX9.7 At Least One Fault or Status Message (DBX0.0...9.3)
  END_STRUCT ;
BEGIN
   Fuse_Fault := FALSE;
   Motor_Protect := FALSE;
   Motor_Temp := FALSE;
   Air_Low := FALSE;
   EStop_Desk_X120 := FALSE;
   EStop_Desk_X121 := FALSE;
   EStop_Elevator := FALSE;
   EStop_Flipper := FALSE;
   Door_Feeder := FALSE;
   Door_Elevator := FALSE;
   Door_Flipper := FALSE;
   Spare_1_3 := FALSE;
   Spare_1_4 := FALSE;
   Spare_1_5 := FALSE;
   Spare_1_6 := FALSE;
   Spare_1_7 := FALSE;
   C2_Angle_Fault := FALSE;
   Elev_Rollers_Fault := FALSE;
   Elev_Pusher_Fault := FALSE;
   Elev_Not_Centered := FALSE;
   C4_Fault := FALSE;
   C4_Timeout := FALSE;
   C4_Infeed_Obstruct := FALSE;
   C6_Fault := FALSE;
   Flipper_Obstruct := FALSE;
   C10_Fault := FALSE;
   Pivot_Timeout := FALSE;
   Pivot_Conflict := FALSE;
   C13_Delivery_Fault := FALSE;
   C23_Delivery_Fault := FALSE;
   Spare_3_6 := FALSE;
   Spare_3_7 := FALSE;
   VFD_U44_3 := FALSE;
   VFD_U45_0 := FALSE;
   VFD_U45_3 := FALSE;
   VFD_U45_6 := FALSE;
   VFD_U46_0 := FALSE;
   VFD_U46_4 := FALSE;
   VFD_U47_0 := FALSE;
   VFD_U47_5 := FALSE;
   VFD_U47_6 := FALSE;
   VFD_U48_0 := FALSE;
   VFD_U48_3 := FALSE;
   VFD_U48_6 := FALSE;
   VFD_U49_0 := FALSE;
   VFD_U53_2 := FALSE;
   VFD_U53_4 := FALSE;
   VFD_U54_0 := FALSE;
   Sens_B5_1_On := FALSE;
   Sens_B5_2_On := FALSE;
   Sens_B5_4_On := FALSE;
   Sens_B5_5_On := FALSE;
   Sens_B6_0_On := FALSE;
   Sens_B6_7_On := FALSE;
   Sens_B7_0_On := FALSE;
   Sens_B7_1_On := FALSE;
   Sens_B7_2_On := FALSE;
   Sens_B7_3_On := FALSE;
   Sens_B7_4_On := FALSE;
   Sens_B8_2_On := FALSE;
   Sens_B9_6_On := FALSE;
   Sens_B9_7_On := FALSE;
   Sens_B10_4_On := FALSE;
   Sens_B10_5_On := FALSE;
   Sens_B10_7_On := FALSE;
   Sens_B11_0_On := FALSE;
   Sens_B11_1_On := FALSE;
   Sens_B5_4_Off := FALSE;
   Sens_B9_7_Off := FALSE;
   Spare_8_5 := FALSE;
   Spare_8_6 := FALSE;
   Spare_8_7 := FALSE;
   Clearing_Active := FALSE;
   Packets_Present := FALSE;
   Control_Off := FALSE;
   Start_Ready := FALSE;
   Spare_9_4 := FALSE;
   Spare_9_5 := FALSE;
   Any_Fault := FALSE;
   Any_Alarm := FALSE;
END_DATA_BLOCK

DATA_BLOCK "HMI_UPDATE"
TITLE =
VERSION : 0.1


  STRUCT
   HMI_GRAPHIC_TOTAL_1 : DWORD ;	//HMI GRAPHIC TOTAL 1
   HMI_GRAPHIC_TOTAL_2 : DWORD ;	//HMI GRAPHIC TOTAL 1
   HMI_FEED_GRAPHIC : DWORD ;	//HMI GRAPHIC FEED TOTAL 1
   HMI_MOTOR_TOTAL_1 : DWORD ;	//HMI MOTOR TOTAL 1
   HMI_ELEVATOR_PROXS : DWORD ;	//HMI ELEVATOR PROXS
   HMI_FLIPPER_PROXS : DWORD ;	//HMI FLIPPER / TURNTABLE PROXS
   HMI_PUSHER_PROXS : DWORD ;	//HMI PUSHER 9 / PIVOT PROXS
   HMI_FEEDER_PROXS : DWORD ;	//HMI FEEDER PROXS
   HMI_SPARE : DWORD ;	//HMI SPARE
   HMI_FEEDER_GRAPHIC : DWORD ;	//HMI FEEDER GRAPHIC
   HMI_MOTOR_GRAPHIC : DWORD ;	//HMI MOTORGRAPHIC
   HMI_MAIN_PAGE_GRAPHIC : DWORD ;	//HMI MAIN SCREEN GRAPHIC
   HMI_SPARE1 : DWORD ;
   HMI_SPARE2 : DWORD ;
   HMI_SPARE3 : DWORD ;
   HMI_SPARE4 : DWORD ;
   HMI_SPARE5 : DWORD ;
   HMI_SPARE6 : DWORD ;
   HMI_SPARE7 : DWORD ;
   HMI_MOTOR_TOTAL1036 : DWORD ;
   HMI_MOTOR_TOTAL1037 : DWORD ;
   HMI_MOTOR_TOTAL1038 : DWORD ;
   HMI_MOTOR_TOTAL1039 : DWORD ;
   HMI_MOTOR_TOTAL10310 : DWORD ;
  END_STRUCT ;
BEGIN
   HMI_GRAPHIC_TOTAL_1 := DW#16#0;
   HMI_GRAPHIC_TOTAL_2 := DW#16#0;
   HMI_FEED_GRAPHIC := DW#16#0;
   HMI_MOTOR_TOTAL_1 := DW#16#0;
   HMI_ELEVATOR_PROXS := DW#16#0;
   HMI_FLIPPER_PROXS := DW#16#0;
   HMI_PUSHER_PROXS := DW#16#0;
   HMI_FEEDER_PROXS := DW#16#0;
   HMI_SPARE := DW#16#0;
   HMI_FEEDER_GRAPHIC := DW#16#0;
   HMI_MOTOR_GRAPHIC := DW#16#0;
   HMI_MAIN_PAGE_GRAPHIC := DW#16#0;
   HMI_SPARE1 := DW#16#0;
   HMI_SPARE2 := DW#16#0;
   HMI_SPARE3 := DW#16#0;
   HMI_SPARE4 := DW#16#0;
   HMI_SPARE5 := DW#16#0;
   HMI_SPARE6 := DW#16#0;
   HMI_SPARE7 := DW#16#0;
   HMI_MOTOR_TOTAL1036 := DW#16#0;
   HMI_MOTOR_TOTAL1037 := DW#16#0;
   HMI_MOTOR_TOTAL1038 := DW#16#0;
   HMI_MOTOR_TOTAL1039 := DW#16#0;
   HMI_MOTOR_TOTAL10310 := DW#16#0;
END_DATA_BLOCK

DATA_BLOCK "PACKET POSITION DB"
TITLE =Packet Positioning - Flipper C7 + Pusher 2 C9 - Stop Time per Lengt
//One stop time per packet length class (15 mm classes, 510 ... > 975 mm).
//Time = belt run after the packet tail leaves B7.4 (step 8N5 -> 8N6, Timer 42).
//Time_ms[class] = 0 -> Default_ms (1500 = as before v1.0).
//v1.1 2026-11-24: HMI packet drawing: Disp_Length_mm (DBW86) + 4 width class
//bits (DBX90.0...90.3, one ON) from the C10 measured width (DB30 Width_mm_Cal).
//v1.2 2026-11-24: + C9 Pusher 2 conveyor (feeder lateral position, Timer 62): one
//time per length class too, Time 0 = "HMI_DB".CONV_9_POS_mS x 10 (as before).
//DBW98 / DBW100 reserved for the flipper drawing (tail / front, later).
//v1.3 2026-11-24: C9 HMI drawing: one packet drawing, 16 copies at 16 lateral
//positions, one shown (C9_Pos_Bits, one bit ON) from the C9 stop time used.
//v1.4 2026-11-24: DB15 symbol renamed "PACKET POSITION DB" (was "FLIPPER POS DB").
VERSION : 1.4


